(* IEC 61131-3 sources: PLC-IsaVODE/PLC-IsaVODE/samples/plc-programs (part 9) *)

(* ---- 663-GEN_RMP.ST ---- *)
FUNCTION D_TRUNC : DINT
  VAR_INPUT
    x : REAL;
  END_VAR

  D_TRUNC := REAL_TO_DINT(X);
  IF X > 0.0 THEN
  	IF DINT_TO_REAL(D_TRUNC) > X THEN D_TRUNC := D_TRUNC - DINT#1; END_IF;
  ELSE
  	IF DINT_TO_REAL(D_TRUNC) < X THEN D_TRUNC := D_TRUNC + DINT#1; END_IF;
  END_IF;
END_FUNCTION

FUNCTION FRACT:REAL
	VAR_INPUT
		X :	REAL;
	END_VAR

	IF ABS(x) < 2.0E9 THEN
		FRACT := x - DINT_TO_REAL(D_TRUNC(x));
	ELSE
		FRACT := 0.0;
	END_IF;
END_FUNCTION

FUNCTION _REAL_TO_DWORD: DWORD

  VAR_INPUT
    X :	REAL;
  END_VAR

  IF REAL_TO_DWORD(0.5) = DWORD#1 THEN
    _REAL_TO_DWORD := REAL_TO_DWORD(x);
  ELSIF X > 0.0 THEN
    _REAL_TO_DWORD := REAL_TO_DWORD(x+0.5);
  ELSIF X < 0.0 THEN
    _REAL_TO_DWORD := REAL_TO_DWORD(x-0.5);
  ELSE
    _REAL_TO_DWORD := DWORD#0;
  END_IF;
END_FUNCTION

FUNCTION _DWORD_TO_REAL:REAL
	VAR_INPUT
		IN :	DWORD;
	END_VAR

	_DWORD_TO_REAL := UDINT_TO_REAL(DWORD_TO_UDINT(IN));

END_FUNCTION

FUNCTION MULTIME:TIME
	VAR_INPUT
		T :	TIME;
		M :	REAL;
	END_VAR

	multime := DWORD_TO_TIME(_REAL_TO_DWORD(_DWORD_TO_REAL(TIME_TO_DWORD(t))*M));
END_FUNCTION

FUNCTION TIME_TO_REAL1:REAL

VAR_INPUT
	X :	TIME;
END_VAR

TIME_TO_REAL1 := UDINT_TO_REAL(DINT_TO_UDINT(TIME_TO_DINT(X)));
END_FUNCTION

FUNCTION MODR : REAL
  VAR_INPUT
    IN : REAL;
    DIVI : REAL;
  END_VAR

  IF divi = 0.0 THEN
  	MODR := 0.0;
  ELSE
  	MODR := in - DINT_TO_REAL(FLOOR2(in / divi)) * divi;
  END_IF;
END_FUNCTION

FUNCTION FLOOR2 : DINT
  VAR_INPUT
    x : REAL;
  END_VAR

  FLOOR2 := REAL_TO_DINT(X);
  IF DINT_TO_REAL(FLOOR2) > X THEN
  	FLOOR2 := FLOOR2 - DINT#1;
  END_IF;
END_FUNCTION

FUNCTION UDINT_TO_TIME2:TIME

	VAR_INPUT
		IN :	UDINT;
	END_VAR

	UDINT_TO_TIME2 := DINT_TO_TIME(UDINT_TO_DINT(IN));

END_FUNCTION

FUNCTION_BLOCK T_PLC_MS_block
	VAR_OUTPUT
		T_PLC_MS :	UDINT;
	END_VAR

	VAR_EXTERNAL
		PLC_TICKS_PER_SEC :	INT;
		PLC_SYS_TICK_CNT :	DINT;
	END_VAR

	VAR
		debug :	BOOL;(*Debug-Mode ON / OFF*)
		N :	INT;(*Debug-Faktor*)
		Offset :	UDINT;(*Debug-Offset*)
		temp :	DWORD := DWORD#1;(*Debug-Offset*)
		mode :	BOOL;(*modus*)
		faktor :	UDINT;(*Systemtakt-Faktor*)
		init :	BOOL;
		v_plc_ticks_per_sec :	UDINT;
		base :	UDINT := UDINT#1000;
	END_VAR

	IF init = FALSE THEN
		v_plc_ticks_per_sec := INT_TO_UDINT(PLC_TICKS_PER_SEC);
		IF v_plc_ticks_per_sec = UDINT#1024 THEN
			faktor := UDINT#1;
			mode := FALSE;
		ELSIF v_plc_ticks_per_sec > UDINT#0 THEN
			IF v_plc_ticks_per_sec <= base THEN
				faktor := base / v_plc_ticks_per_sec;
				mode := FALSE;
			ELSE
				faktor := v_plc_ticks_per_sec / base;
				mode := TRUE;
			END_IF;
		ELSE
			faktor := UDINT#1;
		END_IF;
		init := TRUE;
	END_IF;

	IF mode THEN
		T_PLC_MS := DINT_TO_UDINT(PLC_SYS_TICK_CNT) / faktor;
	ELSE
		T_PLC_MS := DINT_TO_UDINT(PLC_SYS_TICK_CNT) * faktor;
	END_IF;

	IF debug THEN
		T_PLC_MS := (DWORD_TO_UDINT(SHL(UDINT_TO_DWORD(T_PLC_MS),N) OR SHL(temp,N)) - UDINT#1) + Offset;
	END_IF;

END_FUNCTION_BLOCK

FUNCTION_BLOCK GEN_RMP_Block

	VAR_INPUT
		PT :	TIME := T#1s;
		AM :	REAL := REAL#1.0;
		OS :	REAL;
		DL :	REAL;
	END_VAR

	VAR_OUTPUT
		Q :	BOOL;
		OUT :	REAL;
	END_VAR

	VAR
		tx :	TIME;
		last :	TIME;
		init :	BOOL;
		temp :	REAL;
		ltemp :	REAL;
		T_PLC_MS :	T_PLC_MS_Block;
	END_VAR

	T_PLC_MS();
	tx:= UDINT_TO_TIME(T_PLC_MS.T_PLC_MS) - last;
	DL := modR(dl,1.0);
	IF dl < 0.0 THEN dl := 1.0 - dl; END_IF;

	IF NOT init THEN
		init := TRUE;
		last := tx;
		tx := t#0s;
	END_IF;

	IF tx >= pt THEN
		last := last + pt;
		tx := tx - pt;
	END_IF;

	ltemp := temp;
	IF pt > t#0s THEN temp := fract(TIME_TO_REAL1(tx + multime(pt, dl)) / TIME_TO_REAL1(pt)); END_IF;
	out := am * temp + os;

	Q := temp < ltemp;

END_FUNCTION_BLOCK

PROGRAM program0
  VAR
	PT :	TIME := T#1s;
	AM :	REAL := REAL#1.0;
	OS :	REAL;
	DL :	REAL;
	Q :	BOOL;
	OUT :	REAL;
	func_block : GEN_RMP_Block;
  END_VAR
	func_block.PT  :=PT;
	func_block.AM  :=AM;
	func_block.OS  :=OS;
	func_block.DL  :=DL;
	func_block();
	Q := func_block.Q;
	OUT := func_block.OUT;
END_PROGRAM

CONFIGURATION Config0
	VAR_GLOBAL
		PLC_TICKS_PER_SEC :	INT;
		PLC_SYS_TICK_CNT :	DINT;
	END_VAR
	RESOURCE Res0 ON PLC
		TASK task0(INTERVAL := T#20ms,PRIORITY := 0);
		PROGRAM instance0 WITH task0 : program0;
	END_RESOURCE
END_CONFIGURATION

(* ---- 664-T_AVG24.ST ---- *)
TYPE
  oscat_T_AVG24         	  : ARRAY [0..47]   OF INT;
END_TYPE

FUNCTION_BLOCK T_PLC_MS_block
	VAR_OUTPUT
		T_PLC_MS :	UDINT;
	END_VAR

	VAR_EXTERNAL
		PLC_TICKS_PER_SEC :	INT;
		PLC_SYS_TICK_CNT :	DINT;
	END_VAR

	VAR
		debug :	BOOL;(*Debug-Mode ON / OFF*)
		N :	INT;(*Debug-Faktor*)
		Offset :	UDINT;(*Debug-Offset*)
		temp :	DWORD := DWORD#1;(*Debug-Offset*)
		mode :	BOOL;(*modus*)
		faktor :	UDINT;(*Systemtakt-Faktor*)
		init :	BOOL;
		v_plc_ticks_per_sec :	UDINT;
		base :	UDINT := UDINT#1000;
	END_VAR

	IF init = FALSE THEN
		v_plc_ticks_per_sec := INT_TO_UDINT(PLC_TICKS_PER_SEC);
		IF v_plc_ticks_per_sec = UDINT#1024 THEN
			faktor := UDINT#1;
			mode := FALSE;
		ELSIF v_plc_ticks_per_sec > UDINT#0 THEN
			IF v_plc_ticks_per_sec <= base THEN
				faktor := base / v_plc_ticks_per_sec;
				mode := FALSE;
			ELSE
				faktor := v_plc_ticks_per_sec / base;
				mode := TRUE;
			END_IF;
		ELSE
			faktor := UDINT#1;
		END_IF;
		init := TRUE;
	END_IF;

	IF mode THEN
		T_PLC_MS := DINT_TO_UDINT(PLC_SYS_TICK_CNT) / faktor;
	ELSE
		T_PLC_MS := DINT_TO_UDINT(PLC_SYS_TICK_CNT) * faktor;
	END_IF;

	IF debug THEN
		T_PLC_MS := (DWORD_TO_UDINT(SHL(UDINT_TO_DWORD(T_PLC_MS),N) OR SHL(temp,N)) - UDINT#1) + Offset;
	END_IF;

END_FUNCTION_BLOCK

FUNCTION_BLOCK FILTER_I_Block
	VAR_INPUT
		X :	INT;
		T :	TIME;
	END_VAR

	VAR_OUTPUT
		Y :	INT;
	END_VAR

	VAR
		Yi :	DINT;
		last :	UDINT;
		tx :	UDINT;
		init :	BOOL;
		T_PLC_MS :	T_PLC_MS_block;
	END_VAR

	T_PLC_MS();
	tx:= T_PLC_MS.T_PLC_MS;

	IF NOT init OR T = t#0s THEN
		init := TRUE;
		Yi := INT_TO_DINT(X) * DINT#1000;
	ELSE
		Yi := Yi + INT_TO_DINT(X - Y) * UDINT_TO_DINT(tx - last) * DINT#1000 / TIME_TO_DINT(T);
	END_IF;
	last := tx;
	Y := DINT_TO_INT(yi / DINT#1000);

END_FUNCTION_BLOCK

FUNCTION TIME_TO_UDINT2:UDINT
	VAR_INPUT
		X :	TIME;
	END_VAR

	TIME_TO_UDINT2 := DINT_TO_UDINT(TIME_TO_DINT(X));
END_FUNCTION

FUNCTION INC1:INT

	VAR_INPUT
		X :	INT;
		N :	INT;
	END_VAR

	IF X >= N - 1 THEN
		INC1 := 0;
	ELSE
		INC1 := X + 1;
	END_IF;
END_FUNCTION

FUNCTION_BLOCK T_AVG24_Block

	VAR_INPUT
		TS :	INT;
		DTI :	UDINT;
		RST :	BOOL;
		T_FILTER :	TIME := T#10m;
		SCALE :	REAL := 1.0;
		OFS :	REAL;
	END_VAR

	VAR_OUTPUT
		TA :	REAL;
		_TP :	BOOL;
	END_VAR

	VAR_IN_OUT
		T24 :	REAL;
		T24_MAX :	REAL;
		T24_MIN :	REAL;
	END_VAR

	VAR
		samples :	oscat_T_AVG24;
		pos :	INT;
		init :	BOOL;
		sum :	DINT;
		last :	UDINT;
		tmp_maxxx :	INT;
		tmp_min :	INT;
		i :	INT;
		ft1 :	FILTER_I_Block;
	END_VAR

	ft1(X := TS, T := T_FILTER);

	IF rst OR NOT init THEN
		init := TRUE;
		IF T24 = -1000.0 THEN t24 := INT_TO_REAL(ft1.Y) * 0.1; END_IF;
		FOR pos := 0 TO 47 DO
			samples[pos] := REAL_TO_INT(T24 * 10.0);
		END_FOR;
		pos := 0;
		sum := INT_TO_DINT(samples[0]) * DINT#48;
		TA := (INT_TO_REAL(ft1.Y) * 0.1 + OFS) * SCALE;
		T24 := (DINT_TO_REAL(sum) * 0.00208333333333 + OFS) * SCALE;
		_TP := TRUE;
	ELSIF (dti / UDINT#60 MOD UDINT#30) = UDINT#0 AND DTI > last THEN
		last := DTI + TIME_TO_UDINT2(T#1m);
		sum := sum - INT_TO_DINT(samples[pos]);
		samples[pos] := ft1.Y;
		sum := sum + INT_TO_DINT(samples[pos]);
		pos := INC1(pos, 48);
		TA := (INT_TO_REAL(ft1.Y) * 0.1 + OFS) * SCALE;
		T24 := (DINT_TO_REAL(sum) * 0.00208333333333 + OFS) * SCALE;
		tmp_maxxx := -32000;
		tmp_min := 32000;
		FOR i := 0 TO 47 DO
			tmp_maxxx := MAX(tmp_maxxx, samples[i]);
			tmp_min := MIN(tmp_min, samples[i]);
		END_FOR;
		T24_MAX := (INT_TO_REAL(tmp_maxxx) * 0.1 + OFS) * SCALE;
		T24_MIN := (INT_TO_REAL(tmp_min) * 0.1 + OFS) * SCALE;
		_TP := TRUE;
	ELSE
		_TP := FALSE;
	END_IF;

END_FUNCTION_BLOCK

PROGRAM program0
	VAR
		TS :	INT;
		DTI :	UDINT;
		RST :	BOOL;
		T_FILTER :	TIME := T#10m;
		SCALE :	REAL := 1.0;
		OFS :	REAL;
		TA :	REAL;
		_TP :	BOOL;

		func_block : T_AVG24_Block;
	END_VAR
	func_block.TS := TS;
	func_block.DTI := DTI;
	func_block.RST := RST ;
	func_block.T_FILTER := T_FILTER;
	func_block.SCALE := SCALE;
	func_block.OFS := OFS ;

	func_block();
	TA  := func_block.TA;
	_TP  := func_block._TP;

END_PROGRAM

CONFIGURATION Config0
	VAR_GLOBAL
		PLC_TICKS_PER_SEC :	INT;
		PLC_SYS_TICK_CNT :	DINT;
	END_VAR
  	RESOURCE Res0 ON PLC
    	TASK task0(INTERVAL := T#20ms,PRIORITY := 0);
    	PROGRAM instance0 WITH task0 : program0;
  	END_RESOURCE
END_CONFIGURATION

(* ---- 665-TANK_LEVEL.ST ---- *)
FUNCTION_BLOCK TONOF

	VAR_INPUT
		IN :	BOOL;
		T_ON :	TIME;
		T_OFF :	TIME;
	END_VAR

	VAR_OUTPUT
		Q :	BOOL;
	END_VAR

	VAR
		X :	TON;
		old :	BOOL;
		mode :	BOOL;
	END_VAR

	IF IN XOR old THEN
	X(IN := FALSE, PT := SEL_TIME(IN,T_OFF,T_ON));
	mode := IN;
	old := IN;
	END_IF;
	X(IN := TRUE);
	IF X.Q THEN Q := mode;END_IF;

END_FUNCTION_BLOCK

FUNCTION UDINT_TO_TIME2:TIME

	VAR_INPUT
		IN :	UDINT;
	END_VAR

	UDINT_TO_TIME2 := DINT_TO_TIME(UDINT_TO_DINT(IN));

END_FUNCTION

FUNCTION_BLOCK T_PLC_MS_block
	VAR_OUTPUT
		T_PLC_MS :	UDINT;
	END_VAR

	VAR_EXTERNAL
		PLC_TICKS_PER_SEC :	INT;
		PLC_SYS_TICK_CNT :	DINT;
	END_VAR

	VAR
		debug :	BOOL;(*Debug-Mode ON / OFF*)
		N :	INT;(*Debug-Faktor*)
		Offset :	UDINT;(*Debug-Offset*)
		temp :	DWORD := DWORD#1;(*Debug-Offset*)
		mode :	BOOL;(*modus*)
		faktor :	UDINT;(*Systemtakt-Faktor*)
		init :	BOOL;
		v_plc_ticks_per_sec :	UDINT;
		base :	UDINT := UDINT#1000;
	END_VAR

	IF init = FALSE THEN
		v_plc_ticks_per_sec := INT_TO_UDINT(PLC_TICKS_PER_SEC);
		IF v_plc_ticks_per_sec = UDINT#1024 THEN
			faktor := UDINT#1;
			mode := FALSE;
		ELSIF v_plc_ticks_per_sec > UDINT#0 THEN
			IF v_plc_ticks_per_sec <= base THEN
				faktor := base / v_plc_ticks_per_sec;
				mode := FALSE;
			ELSE
				faktor := v_plc_ticks_per_sec / base;
				mode := TRUE;
			END_IF;
		ELSE
			faktor := UDINT#1;
		END_IF;
		init := TRUE;
	END_IF;

	IF mode THEN
		T_PLC_MS := DINT_TO_UDINT(PLC_SYS_TICK_CNT) / faktor;
	ELSE
		T_PLC_MS := DINT_TO_UDINT(PLC_SYS_TICK_CNT) * faktor;
	END_IF;

	IF debug THEN
		T_PLC_MS := (DWORD_TO_UDINT(SHL(UDINT_TO_DWORD(T_PLC_MS),N) OR SHL(temp,N)) - UDINT#1) + Offset;
	END_IF;
END_FUNCTION_BLOCK

FUNCTION TIME_TO_UDINT2:UDINT
	VAR_INPUT
		X :	TIME;
	END_VAR

	TIME_TO_UDINT2 := DINT_TO_UDINT(TIME_TO_DINT(X));
END_FUNCTION

FUNCTION_BLOCK ACTUATOR_COIL_Block

	VAR_INPUT
		IN :	BOOL;
		SELF_ACT_CYCLE :	TIME := T#10d;
		SELF_ACT_TIME :	TIME := T#1s;
	END_VAR

	VAR_OUTPUT
		OUT :	BOOL;
		STATUS :	BYTE;
	END_VAR

	VAR
		last :	UDINT;
		init :	BOOL;
		tx :	UDINT;
		now :	UDINT;
		T_PLC_MS :	T_PLC_MS_Block;
	END_VAR

	T_PLC_MS();
	now := T_PLC_MS.T_PLC_MS;

	IF NOT init THEN
		last := now;
		init := TRUE;
	ELSIF IN THEN
		OUT := TRUE;
		STATUS := BYTE#101;
		LAST := now;
	ELSE
		OUT := FALSE;
		STATUS := BYTE#100;
		tx := now - last;
		IF (self_act_cycle > T#0s) AND (tx >= TIME_TO_UDINT2(self_act_cycle)) THEN
			OUT := TRUE;
			STATUS := BYTE#102;
			IF tx >= TIME_TO_UDINT2(self_act_cycle + self_act_time) THEN
				last := now;
				OUT := FALSE;
				STATUS := BYTE#100;
			END_IF;
		END_IF;
	END_IF;

END_FUNCTION_BLOCK

FUNCTION_BLOCK TANK_LEVEL_Block

	VAR_INPUT
		LEVEL :	BOOL;
		LEAK :	BOOL;
		ACLR :	BOOL;
		MAX_VALVE_TIME :	TIME;
		LEVEL_DELAY_TIME :	TIME;
	END_VAR

	VAR_OUTPUT
		VALVE :	BOOL;
		ALARM :	BOOL;
		STATUS :	BYTE;
	END_VAR

	VAR
		cx :	ACTUATOR_COIL_Block;
		tn :	TON;
		tl :	TONOF;
		open :	BOOL;
	END_VAR

	tl(in := level, T_ON := level_delay_time, T_OFF := level_delay_time);
	open := tl.Q;

	IF ALARM THEN
		IF ACLR THEN
			ALARM := FALSE;
			STATUS := BYTE#101;
			cx(in := FALSE);
		END_IF;
		RETURN;
	ELSIF LEAK THEN
		cx(in := FALSE);
		ALARM := TRUE;
		STATUS := BYTE#1;
	ELSIF open THEN
		cx(in := TRUE);
		STATUS := BYTE#102;
	ELSE
		cx(in := FALSE);
		STATUS := BYTE#100;
	END_IF;

	tn(in := cx.out AND (MAX_VALVE_TIME > T#0s), PT := MAX_VALVE_TIME);
	IF tn.Q THEN
		ALARM := TRUE;
		STATUS := BYTE#2;
		cx(in := FALSE);
	END_IF;

	VALVE := cx.out;
END_FUNCTION_BLOCK

PROGRAM program0
	VAR
		LEVEL :	BOOL;
		LEAK :	BOOL;
		ACLR :	BOOL;
		MAX_VALVE_TIME :	TIME;
		LEVEL_DELAY_TIME :	TIME;
		VALVE :	BOOL;
		ALARM :	BOOL;
		STATUS :	BYTE;

		func_block : TANK_LEVEL_Block;
	END_VAR
	func_block.LEVEL := LEVEL;
	func_block.LEAK := LEAK;
	func_block.ACLR := ACLR ;
	func_block.MAX_VALVE_TIME := MAX_VALVE_TIME;
	func_block.LEVEL_DELAY_TIME := LEVEL_DELAY_TIME ;
	func_block();
	VALVE  := func_block.VALVE;
	ALARM  := func_block.ALARM;
	STATUS  := func_block.STATUS;
END_PROGRAM

CONFIGURATION Config0
	VAR_GLOBAL
		PLC_TICKS_PER_SEC :	INT;
		PLC_SYS_TICK_CNT :	DINT;
	END_VAR
  	RESOURCE Res0 ON PLC
    	TASK task0(INTERVAL := T#20ms,PRIORITY := 0);
    	PROGRAM instance0 WITH task0 : program0;
  	END_RESOURCE
END_CONFIGURATION

(* ---- 666-M_TX.ST ---- *)
FUNCTION_BLOCK T_PLC_MS_block
	VAR_OUTPUT
		T_PLC_MS :	UDINT;
	END_VAR

	VAR_EXTERNAL
		PLC_TICKS_PER_SEC :	INT;
		PLC_SYS_TICK_CNT :	DINT;
	END_VAR

	VAR
		debug :	BOOL;(*Debug-Mode ON / OFF*)
		N :	INT;(*Debug-Faktor*)
		Offset :	UDINT;(*Debug-Offset*)
		temp :	DWORD := DWORD#1;(*Debug-Offset*)
		mode :	BOOL;(*modus*)
		faktor :	UDINT;(*Systemtakt-Faktor*)
		init :	BOOL;
		v_plc_ticks_per_sec :	UDINT;
		base :	UDINT := UDINT#1000;
	END_VAR

	IF init = FALSE THEN
		v_plc_ticks_per_sec := INT_TO_UDINT(PLC_TICKS_PER_SEC);
		IF v_plc_ticks_per_sec = UDINT#1024 THEN
			faktor := UDINT#1;
			mode := FALSE;
		ELSIF v_plc_ticks_per_sec > UDINT#0 THEN
			IF v_plc_ticks_per_sec <= base THEN
				faktor := base / v_plc_ticks_per_sec;
				mode := FALSE;
			ELSE
				faktor := v_plc_ticks_per_sec / base;
				mode := TRUE;
			END_IF;
		ELSE
			faktor := UDINT#1;
		END_IF;
		init := TRUE;
	END_IF;

	IF mode THEN
		T_PLC_MS := DINT_TO_UDINT(PLC_SYS_TICK_CNT) / faktor;
	ELSE
		T_PLC_MS := DINT_TO_UDINT(PLC_SYS_TICK_CNT) * faktor;
	END_IF;

	IF debug THEN
		T_PLC_MS := (DWORD_TO_UDINT(SHL(UDINT_TO_DWORD(T_PLC_MS),N) OR SHL(temp,N)) - UDINT#1) + Offset;
	END_IF;
END_FUNCTION_BLOCK

FUNCTION_BLOCK M_TX_Block

	VAR_INPUT
		IN :	BOOL;
		TMAX :	TIME := t#10d;
		RST :	BOOL;
	END_VAR

	VAR_OUTPUT
		TH :	TIME;
		TL :	TIME;
		DC :	REAL;
		F :	REAL;
		ET :	TIME;
	END_VAR

	VAR
		edge :	BOOL;
		start :	TIME;
		stop :	TIME;
		tx :	TIME;
		rise :	BOOL;
		fall :	BOOL;
		startup :	BOOL;
		T_PLC_MS :	T_PLC_MS_block;
	END_VAR

	IF rst OR (et >= tmax) THEN
		rise := FALSE;
		fall := FALSE;
		startup := FALSE;
		th := t#0ms;
		tl := t#0ms;
		DC := 0.0;
		F := 0.0;
		ET := t#0s;
	END_IF;

	(* avoid timers to start when input is true at startup *)
	IF NOT startup THEN
		edge := in;
		startup := TRUE;
	END_IF;

	(* read system timer *)
	T_PLC_MS();
	tx:= UDINT_TO_TIME(T_PLC_MS.T_PLC_MS);

	(* edge trigger rising and falling edge *)
	IF in XOR edge THEN
		edge := in;
		(* rising edge starts measurement *)
		IF in THEN
			start := Tx;
			rise := TRUE;
			IF fall THEN tl := start - stop; END_IF;
			IF th > t#0ms AND tl > t#0ms THEN
				dc := TIME_TO_REAL(th) / TIME_TO_REAL(th+tl);
				f := 1000.0 / TIME_TO_REAL(th + tl);
			END_IF;
		(* falling edge starts second cycle measurement *)
		ELSE
			stop := Tx;
			fall := TRUE;
			IF rise THEN th := stop - start; END_IF;
			IF th > t#0ms AND tl > t#0ms THEN
				dc := TIME_TO_REAL(th) /  TIME_TO_REAL(th+tl);
				f := 1000.0 / TIME_TO_REAL(th + tl);
			END_IF;
		END_IF;
	END_IF;
	IF rise THEN et := tx - start; END_IF;

	(* check FOR rst input *)
	IF rst OR (et >= tmax) THEN
		rise := FALSE;
		fall := FALSE;
		startup := FALSE;
		th := t#0ms;
		tl := t#0ms;
		DC := 0.0;
		F := 0.0;
		ET := t#0s;
	END_IF;

	(* avoid timers to start when input is true at startup *)
	IF NOT startup THEN
		edge := in;
		startup := TRUE;
	END_IF;

	(* read system timer *)
	T_PLC_MS();
	tx:= UDINT_TO_TIME(T_PLC_MS.T_PLC_MS);

	(* edge trigger rising and falling edge *)
	IF in XOR edge THEN
		edge := in;
		(* rising edge starts measurement *)
		IF in THEN
			start := Tx;
			rise := TRUE;
			IF fall THEN tl := start - stop; END_IF;
			IF th > t#0ms AND tl > t#0ms THEN
				dc := TIME_TO_REAL(th) / TIME_TO_REAL(th+tl);
				f := 1000.0 / TIME_TO_REAL(th + tl);
			END_IF;
		(* falling edge starts second cycle measurement *)
		ELSE
			stop := Tx;
			fall := TRUE;
			IF rise THEN th := stop - start; END_IF;
			IF th > t#0ms AND tl > t#0ms THEN
				dc := TIME_TO_REAL(th) /  TIME_TO_REAL(th+tl);
				f := 1000.0 / TIME_TO_REAL(th + tl);
			END_IF;
		END_IF;
	END_IF;
	IF rise THEN et := tx - start; END_IF;

END_FUNCTION_BLOCK

PROGRAM program0

	VAR
		IN :	BOOL;
		TMAX :	TIME := t#10d;
		RST :	BOOL;

		TH :	TIME;
		TL :	TIME;
		DC :	REAL;
		F :	REAL;
		ET :	TIME;

		func_block : M_TX_Block;
	END_VAR
	func_block.IN := IN;
	func_block.TMAX := TMAX;
	func_block.RST := RST;

	func_block();
	TH := func_block.TH;
	TL := func_block.TL;
	DC := func_block.DC;
	F := func_block.F;
	ET := func_block.ET;

END_PROGRAM

CONFIGURATION Config0

	VAR_GLOBAL
		PLC_TICKS_PER_SEC :	INT;
		PLC_SYS_TICK_CNT :	DINT;
	END_VAR

	RESOURCE Res0 ON PLC
		TASK task0(INTERVAL := T#20ms,PRIORITY := 0);
		PROGRAM instance0 WITH task0 : program0;
	END_RESOURCE

END_CONFIGURATION

(* ---- 667-METER_STAT.ST ---- *)
FUNCTION DAY_OF_WEEK:INT

	VAR_INPUT
		IDATE :	UDINT;
	END_VAR

	DAY_OF_WEEK := UDINT_TO_INT((idate / UDINT#86400 + UDINT#3) MOD UDINT#7) + INT#01;
END_FUNCTION

FUNCTION LEAP_OF_DATE:BOOL

	VAR_INPUT
		IDATE :	UDINT;
	END_VAR

	LEAP_OF_DATE := SHL(UDINT_TO_DWORD((idate + UDINT#43200) / UDINT#31557600), 30) = DWORD#16#80000000;
END_FUNCTION

FUNCTION DAY_OF_YEAR:INT
	VAR_INPUT
		IDATE :	UDINT;
	END_VAR

	DAY_OF_YEAR := UDINT_TO_INT(((idate) / UDINT#86400) MOD UDINT#1461);
	IF DAY_OF_YEAR > 729 THEN
		IF DAY_OF_YEAR > 1095 THEN DAY_OF_YEAR := DAY_OF_YEAR - 1095; ELSE DAY_OF_YEAR := DAY_OF_YEAR - 729; END_IF;
	ELSIF DAY_OF_YEAR > 364 THEN
		DAY_OF_YEAR := DAY_OF_YEAR - 364;
	ELSE
		DAY_OF_YEAR := DAY_OF_YEAR + 1;
	END_IF;
END_FUNCTION

FUNCTION MONTH_OF_DATE:INT

	VAR_INPUT
		IDATE :	UDINT;
	END_VAR

	MONTH_OF_DATE := DAY_OF_YEAR(idate);
	IF MONTH_OF_DATE < 32 THEN
		MONTH_OF_DATE := 1;
	ELSIF LEAP_OF_DATE((IDATE)) THEN
		MONTH_OF_DATE := (MONTH_OF_DATE * 53 + 1668) / 1623;
	ELSE
		MONTH_OF_DATE := (MONTH_OF_DATE * 53 + 1700) / 1620;
	END_IF;
END_FUNCTION

FUNCTION YEAR_OF_DATE:INT
	VAR_INPUT
		IDATE :	UDINT;
	END_VAR

	YEAR_OF_DATE := UDINT_TO_INT((idate+UDINT#43200) / UDINT#31557600 + UDINT#1970);
END_FUNCTION

FUNCTION_BLOCK METER_STAT_Block

	VAR_INPUT
		IN :	REAL;
		DI :	UDINT;
		RST :	BOOL;
	END_VAR

	VAR_IN_OUT
		LAST_DAY :	REAL;
		CURRENT_DAY :	REAL;
		LAST_WEEK :	REAL;
		CURRENT_WEEK :	REAL;
		LAST_MONTH :	REAL;
		CURRENT_MONTH :	REAL;
		LAST_YEAR :	REAL;
		CURRENT_YEAR :	REAL;
	END_VAR

	VAR RETAIN
		year_start :	REAL;
		month_start :	REAL;
		week_start :	REAL;
		day_start :	REAL;
		last_run :	UDINT;
	END_VAR

	IF rst THEN
		Last_Day := 0.0;
		Current_Day := 0.0;
		Day_start := IN;
		Last_week := 0.0;
		Current_week := 0.0;
		Week_start := in;
		Last_month := 0.0;
		Current_month := 0.0;
		month_start := in;
		last_year := 0.0;
		current_year := 0.0;
		year_start := in;
	ELSE
		Current_Day := IN - Day_Start;
		Current_Week := In - Week_Start;
		Current_Month := IN - Month_Start;
		Current_Year := IN - Year_Start;
	END_IF;

	IF YEAR_OF_DATE(DI) > YEAR_OF_DATE(last_run) THEN
		(* a new year has started *)
		last_year := current_year;
		current_year := 0.0;
		year_start := in;
		last_month := current_month;
		current_month := 0.0;
		month_start := in;
		last_day := current_day;
		current_day := 0.0;
		day_start := in;
	ELSIF MONTH_OF_DATE(DI) > MONTH_OF_DATE(last_run) THEN
		(* a new month has started, january is alrerady done by year change *)
		last_month := current_month;
		current_month := 0.0;
		month_start := in;
		last_day := current_day;
		current_day := 0.0;
		day_start := in;
	ELSIF DAY_OF_YEAR(di) > DAY_OF_YEAR(last_run) THEN
		(* day has chaged, first day of year and first day of month has already been taken care of *)
		last_day := current_day;
		current_day := 0.0;
		day_start := in;
	END_IF;
	IF DAY_OF_WEEK(DI) < DAY_OF_WEEK(last_run) THEN
		(* a new week has started *)
		last_week := current_week;
		current_week := 0.0;
		week_start := in;
	END_IF;
	last_run := di;

END_FUNCTION_BLOCK

PROGRAM program0

	VAR
		IN :	REAL;
		DI :	UDINT;
		RST :	BOOL;

		LAST_DAY :	REAL;
		CURRENT_DAY :	REAL;
		LAST_WEEK :	REAL;
		CURRENT_WEEK :	REAL;
		LAST_MONTH :	REAL;
		CURRENT_MONTH :	REAL;
		LAST_YEAR :	REAL;
		CURRENT_YEAR :	REAL;

		func_block : METER_STAT_Block;
	END_VAR

	func_block.IN := IN;
	func_block.DI := DI;
	func_block.RST := RST;
	func_block.LAST_DAY := LAST_DAY;
	func_block.CURRENT_DAY := CURRENT_DAY;
	func_block.LAST_WEEK := LAST_WEEK;
	func_block.CURRENT_WEEK := CURRENT_WEEK;
	func_block.LAST_MONTH := LAST_MONTH;
	func_block.CURRENT_MONTH := CURRENT_MONTH;
	func_block.LAST_YEAR := LAST_YEAR;
	func_block.CURRENT_YEAR := CURRENT_YEAR;

	func_block();

	LAST_DAY  := func_block.LAST_DAY;
	CURRENT_DAY  := func_block.CURRENT_DAY;
	LAST_WEEK  := func_block.LAST_WEEK;
	CURRENT_WEEK  := func_block.CURRENT_WEEK;
	LAST_MONTH  := func_block.LAST_MONTH;
	CURRENT_MONTH  := func_block.CURRENT_MONTH;
	LAST_YEAR  := func_block.LAST_YEAR;
	CURRENT_YEAR  := func_block.CURRENT_YEAR;

END_PROGRAM

CONFIGURATION Config0

	VAR_GLOBAL
		PLC_TICKS_PER_SEC :	INT;
		PLC_SYS_TICK_CNT :	DINT;
	END_VAR

	RESOURCE Res0 ON PLC
		TASK task0(INTERVAL := T#20ms,PRIORITY := 0);
		PROGRAM instance0 WITH task0 : program0;
	END_RESOURCE

END_CONFIGURATION

(* ---- 668-TN_SC_WRITE_C.ST ---- *)
TYPE
  bya_TN_CHAR:       	ARRAY [0..1919] OF BYTE;
  bya_TN_BACKUP:     	ARRAY [0..1919] OF BYTE;
  bya_TN_COLOR:      	ARRAY [0..1919] OF BYTE;
  bya_TN_Line_Update:	ARRAY [0..23]   OF BOOL;

  us_TN_SCREEN :
  STRUCT
		bya_CHAR:			bya_TN_CHAR;
		bya_COLOR:			bya_TN_COLOR;
		bya_BACKUP:			bya_TN_BACKUP;
		bya_Line_Update:	bya_TN_Line_Update;

		by_Input_Exten_Code:    BYTE;
		by_Input_ASCII_Code:    BYTE;
		bo_Input_ASCII_IsNum:   BOOL;
		in_Page_Number:        	INT;                (* aktive Seiten-Nr.              *)
		in_Cursor_X:           	INT;                (* Cursor X-Position              *)
		in_Cursor_Y:           	INT;                (* Cursor Y-Position              *)
		in_EOS_Offset:         	INT;                (* End of String Offset           *)
		by_Clear_Screen_Attr:  	BYTE;               (* Clear-Screen Attr              *)
		bo_Clear_Screen:       	BOOL;               (* Clear-Screen ausl�sen          *)
		bo_Modal_Dialog:       	BOOL;               (* Modaler Dialog ist aktiv       *)
		bo_Menue_Bar_Dialog:   	BOOL;               (* Menue Dialog ist aktiv         *)

  END_STRUCT;
END_TYPE

FUNCTION _BYTE_TO_INT:INT
	VAR_INPUT
		IN :	BYTE;
	END_VAR

	_BYTE_TO_INT := USINT_TO_INT(BYTE_TO_USINT(IN));
END_FUNCTION

FUNCTION_BLOCK CHR_TO_STRING_Block
	VAR_INPUT
		C :	BYTE;
	END_VAR

	VAR_OUTPUT
		CHR_TO_STRING :	STRING;
	END_VAR

	CHR_TO_STRING := BYTE_TO_STRING(C);

END_FUNCTION_BLOCK

FUNCTION BIT_OF_DWORD : BOOL
  VAR_INPUT
    IN : DWORD;
    N : INT;
  END_VAR

  BIT_OF_DWORD := (SHR(in,N) AND 16#00000001) > 0;
  (* from OSCAT library; www.oscat.de  *)
END_FUNCTION

FUNCTION_BLOCK FILL_Block
	VAR_INPUT
		C :	BYTE;
		L :	INT;
	END_VAR

	VAR_OUTPUT
		FILL :	STRING;
	END_VAR

	VAR
		N :	BYTE;
		I :	INT;
		sx :	STRING;
		CHR_TO_STRING :	CHR_TO_STRING_Block;
		FILL_tmp :	STRING;
	END_VAR

	CHR_TO_STRING(C:=c);
	Sx:=CHR_TO_STRING.CHR_TO_STRING;
	(* create string *)
	N := INT_TO_BYTE(LIMIT(0,L,80));
	(* create a string of characters to be connected to str *)
	FILL := '';
	FOR i := 1 TO 8 DO
		FILL_tmp := FILL;
		FILL := CONCAT(FILL_tmp,FILL);
		IF BIT_OF_DWORD(BYTE_TO_DWORD(N),7) THEN FILL := CONCAT(FILL,Sx); END_IF;
		N := SHL(N,1);
	END_FOR;
END_FUNCTION_BLOCK

FUNCTION_BLOCK FIX_Block

	VAR_INPUT
		STR :	STRING;
		L :	INT;
		C :	BYTE;
		M :	INT;
	END_VAR

	VAR_OUTPUT
		FIX :	STRING;
	END_VAR

	VAR
		N :	INT;
		FILL :	FILL_Block;
	END_VAR

	N := LIMIT(0,L,255) - LEN(str);
	IF N <= 0 THEN
		(* truncate the string at length N *)
		IF M = 1 THEN
			FIX := RIGHT(str,L);
		ELSE
			FIX := LEFT(str,L);
		END_IF;
	ELSIF M = 1 THEN
		(* connect fill characters at the beginning *)
		FILL(C:=C,L:=N);
		FIX := CONCAT(FILL.FILL,str);
	ELSIF M = 2 THEN
		(* center str beween fill characters *)
		(* for an uneven number of fill characters, there is one more at the end *)
		FILL(C:=C,L:=_BYTE_TO_INT(SHR(INT_TO_BYTE(N+1),1)));
		FIX := CONCAT(str,FILL.FILL);
		FILL(C:=C,L:=_BYTE_TO_INT(SHR(INT_TO_BYTE(N),1)));
		FIX := CONCAT(FILL.FILL,FIX);
	ELSE
		(* connect fill characters at the end *)
		FILL(C:=C,L:=N);
		FIX := CONCAT(str,FILL.FILL);
	END_IF;

END_FUNCTION_BLOCK

FUNCTION_BLOCK TN_SC_WRITE_C_Block

	VAR
		FB_FIX :	FIX_Block;
		FB_TN_SC_WRITE :	TN_SC_WRITE;
	END_VAR

	VAR_INPUT
		Iin_Y :	INT;
		Iin_X :	INT;
		Iby_ATTR :	BYTE;
		Ist_STRING :	STRING;
		Iin_LENGTH :	INT;
		Iin_OPTION :	INT;
	END_VAR

	VAR_IN_OUT
		Xus_TN_SCREEN :	us_TN_SCREEN;
	END_VAR

	FB_FIX.str:=Ist_STRING;
	FB_FIX.L:=Iin_LENGTH;
	FB_FIX.C:=BYTE#32;
	FB_FIX.M:=Iin_OPTION;
	FB_FIX();

	FB_TN_SC_WRITE.Iin_Y			:= Iin_Y;
	FB_TN_SC_WRITE.Iin_X			:= Iin_X;
	FB_TN_SC_WRITE.Iby_ATTR			:= Iby_ATTR;
	FB_TN_SC_WRITE.Ist_STRING		:= FB_FIX.FIX;
	FB_TN_SC_WRITE.Xus_TN_SCREEN	:= Xus_TN_SCREEN;
	FB_TN_SC_WRITE();
	Xus_TN_SCREEN := FB_TN_SC_WRITE.Xus_TN_SCREEN;

END_FUNCTION_BLOCK

PROGRAM program0
	VAR
		Iin_Y :	INT;
		Iin_X :	INT;
		Iby_CHAR :	BYTE;
		Xus_TN_SCREEN :	us_TN_SCREEN;

		func_block : TN_SC_WRITE_C_Block;
	END_VAR
	func_block.Iin_Y := Iin_Y;
	func_block.Iin_X := Iin_X;
	func_block.Iby_CHAR := Iby_CHAR;
	func_block.Xus_TN_SCREEN := Xus_TN_SCREEN;

	func_block();
	Xus_TN_SCREEN  := func_block.Xus_TN_SCREEN;
END_PROGRAM

CONFIGURATION Config0
	RESOURCE Res0 ON PLC
		TASK task0(INTERVAL := T#20ms,PRIORITY := 0);
		PROGRAM instance0 WITH task0 : program0;
	END_RESOURCE
END_CONFIGURATION

(* ---- 669-MONTH_TO_STRING.ST ---- *)
TYPE
  oscat_ELEMENT_MONTHS 	: ARRAY [1..12] OF STRING;
  oscat_MONTHS			: ARRAY [1..3]  OF oscat_ELEMENT_MONTHS := [0, 0, 0];
  oscat_ELEMENT_MONTHS3	: ARRAY [1..12] OF STRING;
  oscat_MONTHS3			: ARRAY [1..3]  OF oscat_ELEMENT_MONTHS3 := [0,0,0];
END_TYPE

TYPE oscat_LANGUAGE:
  STRUCT
    DEFAULT 	: INT;
	LMAX    	: INT;
  END_STRUCT;
END_TYPE

FUNCTION_BLOCK SETUP_LANGUAGE_Block

	VAR_IN_OUT
		LANGUAGE :	oscat_LANGUAGE;
	END_VAR

	VAR
		init :	BOOL;
	END_VAR

	IF init THEN RETURN; END_IF;
	init := TRUE;

	LANGUAGE.DEFAULT  := 1; (* 1=english, 2=german 3=french *)
	LANGUAGE.LMAX := 3;
END_FUNCTION_BLOCK

FUNCTION_BLOCK SETUP_MONTHS3_Block

	VAR_IN_OUT
		MONTHS3 :	oscat_MONTHS3;
	END_VAR

	VAR
		init :	BOOL;
	END_VAR

	IF init THEN RETURN; END_IF;
	init := TRUE;

	(* ---- english --- *)
	MONTHS3[1][01] := 'Jan';
	MONTHS3[1][02] := 'Feb';
	MONTHS3[1][03] := 'Mar';
	MONTHS3[1][04] := 'Apr';
	MONTHS3[1][05] := 'May';
	MONTHS3[1][06] := 'Jun';
	MONTHS3[1][07] := 'Jul';
	MONTHS3[1][08] := 'Aug';
	MONTHS3[1][09] := 'Sep';
	MONTHS3[1][10] := 'Oct';
	MONTHS3[1][11] := 'Nov';
	MONTHS3[1][12] := 'Dec';

	(* ---- german --- *)
	MONTHS3[2][01] := 'Jan';
	MONTHS3[2][02] := 'Feb';
	MONTHS3[2][03] := 'Mrz';
	MONTHS3[2][04] := 'Apr';
	MONTHs3[2][05] := 'Mai';
	MONTHS3[2][06] := 'Jun';
	MONTHS3[2][07] := 'Jul';
	MONTHS3[2][08] := 'Aug';
	MONTHS3[2][09] := 'Sep';
	MONTHS3[2][10] := 'Okt';
	MONTHS3[2][11] := 'Nov';
	MONTHS3[2][12] := 'Dez';

	(* ---- french --- *)
	MONTHS3[3][01] := 'Jan';
	MONTHS3[3][02] := 'Fev';
	MONTHS3[3][03] := 'Mar';
	MONTHS3[3][04] := 'Avr';
	MONTHs3[3][05] := 'Mai';
	MONTHS3[3][06] := 'Jun';
	MONTHS3[3][07] := 'Jul';
	MONTHS3[3][08] := 'Aou';
	MONTHS3[3][09] := 'Sep';
	MONTHS3[3][10] := 'Oct';
	MONTHS3[3][11] := 'Nov';
	MONTHS3[3][12] := 'Dec';
	(*@KEY@: END_WORKSHEET *)
END_FUNCTION_BLOCK

FUNCTION_BLOCK SETUP_MONTHS_Block

	VAR_IN_OUT
		MONTHS :	oscat_MONTHS;
	END_VAR

	VAR
		init :	BOOL;
	END_VAR

	IF init THEN RETURN; END_IF;
	init := TRUE;

	(* ---- english --- *)
	MONTHS[1][01] := 'January';
	MONTHS[1][02] := 'February';
	MONTHS[1][03] := 'March';
	MONTHS[1][04] := 'April';
	MONTHS[1][05] := 'May';
	MONTHS[1][06] := 'June';
	MONTHS[1][07] := 'July';
	MONTHS[1][08] := 'August';
	MONTHS[1][09] := 'September';
	MONTHS[1][10] := 'October';
	MONTHS[1][11] := 'November';
	MONTHS[1][12] := 'December';

	(* ---- german --- *)
	MONTHS[2][01] := 'Januar';
	MONTHS[2][02] := 'Februar';
	MONTHS[2][03] := 'March';
	MONTHS[2][04] := 'April';
	MONTHS[2][05] := 'Mai';
	MONTHS[2][06] := 'Juni';
	MONTHS[2][07] := 'Juli';
	MONTHS[2][08] := 'August';
	MONTHS[2][09] := 'September';
	MONTHS[2][10] := 'Oktober';
	MONTHS[2][11] := 'November';
	MONTHS[2][12] := 'Dezember';

	(* ---- french --- *)
	MONTHS[3][01] := 'Janvier';
	MONTHS[3][02] := 'Fvrier';
	MONTHS[3][03] := 'mars';
	MONTHS[3][04] := 'Avril';
	MONTHS[3][05] := 'Mai';
	MONTHS[3][06] := 'Juin';
	MONTHS[3][07] := 'Juillet';
	MONTHS[3][08] := 'Aot';
	MONTHS[3][09] := 'Septembre';
	MONTHS[3][10] := 'Octobre';
	MONTHS[3][11] := 'Novembre';
	MONTHS[3][12] := 'Decembre';
END_FUNCTION_BLOCK

FUNCTION_BLOCK MONTH_TO_STRING_Block

	VAR_INPUT
		MTH :	INT;
		LANG :	INT;
		LX :	INT;
	END_VAR

	VAR_OUTPUT
		MONTH_TO_STRING :	STRING;
	END_VAR

	VAR
		LY :	INT;
		SETUP_MONTHS :	SETUP_MONTHS_Block;
		MONTHS :	oscat_MONTHS;
		SETUP_MONTHS3 :	SETUP_MONTHS3_Block;
		MONTHS3 :	oscat_MONTHS3;
		SETUP_LANGUAGE :	SETUP_LANGUAGE_Block;
		LANGUAGE :	oscat_LANGUAGE;
	END_VAR

	SETUP_MONTHS(MONTHS:=MONTHS);
	MONTHS:=SETUP_MONTHS.MONTHS;
	SETUP_MONTHS3(MONTHS3:=MONTHS3);
	MONTHS3:=SETUP_MONTHS3.MONTHS3;
	SETUP_LANGUAGE(LANGUAGE:=LANGUAGE);
	LANGUAGE:=SETUP_LANGUAGE.LANGUAGE;

	IF LANG = 0 THEN Ly := LANGUAGE.DEFAULT; ELSE ly := MIN(LANG, language.LMAX); END_IF;
	IF MTH < 1 OR MTH > 12 THEN
		RETURN;
	ELSIF LX = 0 THEN
		MONTH_TO_STRING := MONTHS[ly][MTH];
	ELSIF Lx = 3 THEN
		MONTH_TO_STRING := MONTHS3[ly][MTH];
	END_IF;

END_FUNCTION_BLOCK

PROGRAM program0
	VAR
		MTH :	INT;
		LANG :	INT;
		LX :	INT;
		MONTH_TO_STRING :	STRING;
		func_block : MONTH_TO_STRING_Block;
	END_VAR
		func_block.MTH  := MTH;
		func_block.LANG  := LANG;
		func_block.LX  := LX;
		func_block();
		MONTH_TO_STRING := func_block.MONTH_TO_STRING;
END_PROGRAM

CONFIGURATION Config0
	RESOURCE Res0 ON PLC
		TASK task0(INTERVAL := T#20ms,PRIORITY := 0);
		PROGRAM instance0 WITH task0 : program0;
	END_RESOURCE
END_CONFIGURATION

(* ---- 670-WORLD_WEATHER_DESC_GE.ST ---- *)
TYPE
  oscat_STRING3               : STRING;
  oscat_STRING8               : STRING;
  oscat_STRING10              : STRING;
  oscat_STRING60              : STRING;
END_TYPE

TYPE
	oscat_WORLD_WEATHER_CUR :
	STRUCT
		OBSERVATION_TIME : oscat_STRING8;
		TEMP_C           : INT;
		WEATHER_CODE     : INT;
		WEATHER_DESC 	 : oscat_STRING60;
		WEATHER_ICON     : INT;
		WIND_SPEED_MILES : INT;
		WIND_SPEED_KMPH  : INT;
		WIND_DIR_DEGREE  : INT;
		WIND_DIR16POINT  : oscat_STRING3;
		PRECIPMM         : REAL;
		HUMIDITY         : INT;
		VISIBILITY       : INT;
		PRESSURE         : INT;
		CLOUDOVER        : INT;
	END_STRUCT;

	oscat_WORLD_WEATHER_DAY :
	STRUCT
		DATE_OF_DAY      : oscat_STRING10;
		TEMP_MAX_C       : INT;
		TEMP_MAX_F       : INT;
		TEMP_MIN_C       : INT;
		TEMP_MIN_F       : INT;
		WIND_SPEED_MILES : INT;
		WIND_SPEED_KMPH  : INT;
		WIND_DIR_DEGREE  : INT;
		WIND_DIR16POINT  : oscat_STRING3;
		WEATHER_CODE     : INT;
		WEATHER_DESC     : oscat_STRING60;
		WEATHER_ICON     : INT;
		PRECIPMM         : REAL;
	END_STRUCT;

	oscat_WORLD_WEATHER_DAY_ARR : ARRAY [0..4] OF oscat_WORLD_WEATHER_DAY;

	oscat_WORLD_WEATHER_DATA :
	STRUCT
		CUR : oscat_WORLD_WEATHER_CUR;
		DAY : oscat_WORLD_WEATHER_DAY_ARR;
	END_STRUCT;

	oscat_WORLD_WEATHER_aI0_41 : ARRAY[0..41] OF INT;
END_TYPE

FUNCTION_BLOCK WORLD_WEATHER_DESC_GE_Block

	VAR_INPUT
		ACTIVATE :	BOOL;
	END_VAR

	VAR_IN_OUT
		WW :	oscat_WORLD_WEATHER_DATA;
	END_VAR

	VAR
		act_last :	BOOL;
		x :	INT;
		y :	INT;
		str :	oscat_STRING60;
		i :	INT;
	END_VAR

	IF ACTIVATE AND act_last = FALSE THEN
		i := 0;
		FOR y := 1 TO 12 DO
			CASE y OF
			1,3,5,7,9:	x :=  WW.DAY[i].WEATHER_CODE;
			2,4,6,8,10:	WW.DAY[i].WEATHER_DESC := str;
						i := i + 1;
			11:			x :=  WW.CUR.WEATHER_CODE;
			12:			WW.CUR.WEATHER_DESC := str;
			END_CASE;

			CASE x OF
				113	:	str := 'heiter/sonnig';
				116	:	str := 'stellenweise wolkig';
				119	:	str := 'wolkig';
				122	:	str := 'awret';
				143	:	str := 'Nebel';
				176	:	str := 'stellenweise nahegelegener Regen';
				179	:	str := 'stellenweise nahegelegener Schneefall';
				182	:	str := 'stellenweise nahegelegener Eisregen';
				185	:	str := 'stellenweise gefrierender Niesel';
				200	:	str := 'nahegelegene Sturm';
				227	:	str := 'Schneetreiben';
				230	:	str := 'Schneesturm';
				248	:	str := 'Nebel';
				260	:	str := 'gefrierender Nebel';
				263	:	str := 'stellenweise leichter Nieselregen';
				266	:	str := 'leichter Niesel';
				281	:	str := 'gefrierender Nieselregen';
				284	:	str := 'stark gefrierender Nieselregen';
				293	:	str := 'stellenweise leichter Regen';
				296	:	str := 'leichter Regen';
				299	:	str := 'zeitweise etwas Regen';
				302	:	str := 'awerg Regen';
				305	:	str := 'zeitweise etwas starker Regen';
				308	:	str := 'starker Regen';
				311	:	str := 'leichter gefrierender Regen';
				314	:	str := 'awerawer oder starker Eisregen';
				317	:	str := 'leichter Eisregen';
				320	:	str := 'awewea oder starker Eisregen';
				323	:	str := 'stellenweise leichter Schneefall';
				326	:	str := 'leichter Scheefall';
				329	:	str := 'stellenweise moderater Schneefall';
				332	:	str := 'awertwy Schnee';
				335	:	str := 'stellenweise starker Scheefall';
				338	:	str := 'starker Schneefall';
				350	:	str := 'Hagel';
				353	:	str := 'leichte ewruerh';
				356	:	str := 'awerwaer oder starker Regenfall';
				359	:	str := 'sintflutartige aweheawh';
				362	:	str := 'leichter Eisregen';
				365	:	str := 'aweraweb oder starker Eisregen';
				368	:	str := 'leichte Schneeschauer';
				371	:	str := 'awerawb oder starker Schneefall';
				374	:	str := 'leichter Hagel';
				377	:	str := 'awerawer oder starker Hagel';
				386	:	str := 'stellenweise leichter Regen in Gewittergebiet';
				389	:	str := 'awer oder starker Regen in Gewittergebiet';
				392	:	str := 'stellenweise leichter Schneefall in Gewittergebiet';
				395	:	str := 'awerh oder starker Schnee in Gewittergebiet';
			ELSE
				str := 	'nicht aweh';
			END_CASE;
		END_FOR;
	END_IF;
	act_last := ACTIVATE;

END_FUNCTION_BLOCK

PROGRAM program0
	VAR
		ACTIVATE :	BOOL;
		WW :	oscat_WORLD_WEATHER_DATA;

		func_block : WORLD_WEATHER_DESC_GE_Block;
	END_VAR
	func_block.ACTIVATE := ACTIVATE;
	func_block.WW := WW;

	func_block();
	WW  := func_block.WW;
END_PROGRAM

CONFIGURATION Config0
	RESOURCE Res0 ON PLC
		TASK task0(INTERVAL := T#20ms,PRIORITY := 0);
		PROGRAM instance0 WITH task0 : program0;
	END_RESOURCE
END_CONFIGURATION

(* ---- 671-LOG_VIEWPORT.ST ---- *)
TYPE
  oscat_STRING80             : STRING;
  oscat_STRING250             : STRING;
END_TYPE

TYPE
  PRINTF_DATA_250  	:  ARRAY [1..11]  OF oscat_STRING250;
  PRINTF_DATA_80 	:  ARRAY [1..11]  OF oscat_STRING80;
  LOG_250       	:  ARRAY [0..400] OF oscat_STRING250;
  LOG_80    		:  ARRAY [0..400] OF oscat_STRING80;
  LOG_OPTION		:  ARRAY [0..400] OF DWORD;

  us_LOG_CONTROL :
  STRUCT
    NEW_MSG              : oscat_STRING250;    (*W neue Nachricht f�r den Datenbuffer   *)
	NEW_MSG_OPTION 		 : DWORD;
    LEVEL                : BYTE;
	SIZE                 : INT;                (*R Anzahl der Strings im LOG_DATA       *)
	RESET                : BOOL;               (*W Nachrichtenbuffer l�schen            *)
    PRINTF               : PRINTF_DATA_250;    (*W Array PRINTF Parameter               *)
    MSG                  : LOG_250;            (*I Array Message                        *)
    MSG_OPTION           : LOG_OPTION;     	   (*I Array Message Option                 *)
	UPDATE_COUNT         : UINT;               (*R Updatez�hler                         *)
    IDX                  : INT;                (*R aktueller Nachrichten-Index          *)
	RING_MODE            : BOOL;               (*I Buffer�berlauf erkannt               *)
  END_STRUCT;

  us_LOG_CONTROL_80 :
  STRUCT
    NEW_MSG              : oscat_STRING80;     (*W neue Nachricht f�r den Datenbuffer   *)
	NEW_MSG_OPTION 		 : DWORD;
    LEVEL                : BYTE;
	SIZE                 : INT;                (*R Anzahl der Strings im LOG_DATA       *)
	RESET                : BOOL;               (*W Nachrichtenbuffer l�schen            *)
    PRINTF               : PRINTF_DATA_80;     (*W Array PRINTF Parameter               *)
    MSG                  : LOG_80;             (*I Array Message                        *)
    MSG_OPTION           : LOG_OPTION;     	   (*I Array Message Option                 *)
	UPDATE_COUNT         : UINT;               (*R Updatez�hler                         *)
    IDX                  : INT;                (*R aktueller Nachrichten-Index          *)
	RING_MODE            : BOOL;               (*I Buffer�berlauf erkannt               *)
  END_STRUCT;

  LINE_ARRAY 			: ARRAY [1..40] OF INT;

  us_LOG_VIEWPORT :
    STRUCT
     LINE_ARRAY          : LINE_ARRAY;
     COUNT               : INT;                (* Anzahl der sichtbaren Nachtrichten   *)
	 UPDATE_COUNT        : UINT;               (* Updatez�hler                         *)
     MOVE_TO_X           : INT;                (* Steuerung der Nachrichtenanzeige     *)
     UPDATE              : BOOL;               (* Daten wurden ge�ndert -> neuzeichnen *)
  END_STRUCT;

END_TYPE

FUNCTION_BLOCK LOG_VIEWPORT_Block

  VAR_IN_OUT
    LC :	us_LOG_CONTROL_80;
    LV :	us_LOG_VIEWPORT;
  END_VAR

  VAR
    pos :	INT;
    count :	INT;
    idx :	INT;
    base :	INT;
    update_pos :	BOOL;
  END_VAR

  IF LV.MOVE_TO_X <> 0 THEN
    CASE LV.MOVE_TO_X OF
    30000:
      pos := 1 ;
    30001:
      pos := LC.SIZE;
    30002:
      pos := pos + LV.COUNT;
    30003:
      pos := pos - LV.COUNT;
    ELSE
      pos := pos + LV.MOVE_TO_X;
    END_CASE;
    update_pos := TRUE;
    LV.MOVE_TO_X := 0;
  END_IF;

  IF (LV.UPDATE_COUNT <> LC.UPDATE_COUNT) OR update_pos THEN
    LV.UPDATE := TRUE;
    LV.UPDATE_COUNT := LC.UPDATE_COUNT;
    update_pos := FALSE;

    IF LC.RING_MODE THEN
      pos := LIMIT(1,pos,LC.SIZE - LV.COUNT + 1);
    ELSE
      IF LC.IDX > LV.COUNT THEN
        pos := LIMIT(1,pos,LC.IDX - LV.COUNT + 1);
      ELSE
        pos := 1;
      END_IF;
    END_IF;

    base := LC.IDX - pos - LV.COUNT + 1;
    IF LC.RING_MODE THEN
      FOR count:= 1 TO LV.COUNT DO
        idx := base + count;
        IF idx < 1 THEN
          idx := idx + LC.SIZE;
        END_IF;
      END_FOR;
    ELSE
      FOR count:= 1 TO LV.COUNT DO
        idx := base + count;
        IF idx < 1 THEN
          LV.LINE_ARRAY[count] := 0;
        ELSE
          LV.LINE_ARRAY[count] := idx;
        END_IF;
      END_FOR;
    END_IF;
  END_IF;

END_FUNCTION_BLOCK

PROGRAM program0
	VAR
		LC :	us_LOG_CONTROL_80;
    LV :	us_LOG_VIEWPORT;

		func_block : LOG_VIEWPORT_Block;
	END_VAR
	func_block.LC := LC;
	func_block.LV := LV;

	func_block();
  LC  := func_block.LC;
  LV  := func_block.LV;

END_PROGRAM

CONFIGURATION Config0

  	RESOURCE Res0 ON PLC
    	TASK task0(INTERVAL := T#20ms,PRIORITY := 0);
    	PROGRAM instance0 WITH task0 : program0;
  	END_RESOURCE

END_CONFIGURATION

(* ---- 672-CTRL_PI.ST ---- *)
FUNCTION_BLOCK T_PLC_US_Block
	VAR_OUTPUT
		T_PLC_US :	UDINT;
	END_VAR

	VAR_EXTERNAL
		PLC_TICKS_PER_SEC :	INT;
		PLC_SYS_TICK_CNT :	DINT;
	END_VAR

	VAR
		debug :	BOOL;
		N :	INT;
		Offset :	UDINT;
		temp :	DWORD := DWORD#1;
		mode :	BOOL;
		faktor :	UDINT;
		init :	BOOL;
		v_plc_ticks_per_sec :	UDINT;
		base :	UDINT := UDINT#1000000;
	END_VAR

	IF init = FALSE THEN
		v_plc_ticks_per_sec := INT_TO_UDINT(PLC_TICKS_PER_SEC);
		IF v_plc_ticks_per_sec = UDINT#1024 THEN
			faktor := UDINT#1000;
			mode := FALSE;
		ELSIF v_plc_ticks_per_sec > UDINT#0 THEN
			IF v_plc_ticks_per_sec <= base THEN
				faktor := base / v_plc_ticks_per_sec;
				mode := FALSE;
			ELSE
				faktor := v_plc_ticks_per_sec / base;
				mode := TRUE;
			END_IF;
		ELSE
			faktor := UDINT#1;
		END_IF;
		init := TRUE;
	END_IF;

	IF mode THEN
		T_PLC_US := DINT_TO_UDINT(PLC_SYS_TICK_CNT) / faktor;
	ELSE
		T_PLC_US := DINT_TO_UDINT(PLC_SYS_TICK_CNT) * faktor;
	END_IF;

	IF debug THEN
		T_PLC_US := (DWORD_TO_UDINT(SHL(UDINT_TO_DWORD(T_PLC_US),N) OR SHL(temp,N)) - UDINT#1) + Offset;
	END_IF;
END_FUNCTION_BLOCK

FUNCTION_BLOCK FT_PIWL

	VAR_INPUT
		IN :	REAL;
		KP :	REAL := 1.0;
		KI :	REAL := 1.0;
		LIM_L :	REAL := -1.0E38;
		LIM_H :	REAL := 1.0E38;
		RST :	BOOL;
	END_VAR

	VAR_OUTPUT
		Y :	REAL;
		LIM :	BOOL;
	END_VAR

	VAR
		init :	BOOL;
		tx :	UDINT;
		tc :	REAL;
		t_last :	UDINT;
		in_last :	REAL;
		i :	REAL;
		p :	REAL;
		T_PLC_US :	T_PLC_US_Block;
	END_VAR

	IF NOT init OR RST THEN
		init := TRUE;
		in_last := in;
		T_PLC_US();
		t_last := T_PLC_US.T_PLC_US;
		i := 0.0;
		tc := 0.0;
	ELSE
		(* read last cycle time in Microseconds *)
		T_PLC_US();
		tx := T_PLC_US.T_PLC_US;
		tc := UDINT_TO_REAL(tx - t_last);
		t_last := tx;

		(* calculate proportional part *)
		p := KP * IN;

		(* run integrator *)
		i := (IN + in_last) * 5.0E-7 * KI * tc + i;
		in_last := IN;

		(* calculate output Y *)
		Y := p + i;

		(* check output for limits *)
		IF Y >= LIM_H THEN
			Y := LIM_H;
			IF ki <> 0.0 THEN
				i := LIM_H - p;
			ELSE
				i := 0.0;
			END_IF;
			LIM := TRUE;
		ELSIF Y <= LIM_L THEN
			Y := LIM_L;
			IF ki <> 0.0 THEN
				i := LIM_L - p;
			ELSE
				i := 0.0;
			END_IF;
			LIM := TRUE;
		ELSE
			LIM := FALSE;
		END_IF;
	END_IF;
END_FUNCTION_BLOCK

FUNCTION_BLOCK CTRL_OUT
	VAR_INPUT
		CI :	REAL;
		OFFSET :	REAL;
		MAN_IN :	REAL;
		LIM_L :	REAL;
		LIM_H :	REAL;
		MANUAL :	BOOL;
	END_VAR

	VAR_OUTPUT
		Y :	REAL;
		LIM :	BOOL;
	END_VAR

	Y := SEL(manual, CI, MAN_IN) + OFFSET;

	IF Y >= LIM_H THEN
		Y := LIM_H;
		LIM := TRUE;
	ELSIF Y <= lim_L THEN
		Y := LIM_L;
		LIM := TRUE;
	ELSE
		LIM := FALSE;
	END_IF;
END_FUNCTION_BLOCK

FUNCTION DEAD_ZONE:REAL

	VAR_INPUT
		X :	REAL;
		L :	REAL;
	END_VAR

	IF ABS(x) > L THEN
		dead_zone := X;
	ELSE
		DEAD_ZONE := 0.0;
	END_IF;

END_FUNCTION

FUNCTION CTRL_IN:REAL
	VAR_INPUT
		SET_POINT :	REAL;
		ACTUAL :	REAL;
		NOISE :	REAL;
	END_VAR
	CTRL_IN := DEAD_ZONE(SET_POINT - ACTUAL, NOISE);
END_FUNCTION

FUNCTION_BLOCK CTRL_PI
	VAR_INPUT
		ACT :	REAL;
		SET :	REAL;
		SUP :	REAL;
		OFS :	REAL;
		M_I :	REAL;
		MAN :	BOOL;
		RST :	BOOL := FALSE;
		KP  :	REAL := 1.0;
		KI  :	REAL := 1.0;
		LL  :	REAL := -1000.0;
		LH  :	REAL := 1000.0;
	END_VAR

	VAR_OUTPUT
		Y    :	REAL;
		DIFF :	REAL;
		LIM  :	BOOL;
	END_VAR

	VAR
		pi :	FT_PIWL;
		co :	CTRL_OUT;
	END_VAR

	DIFF := CTRL_IN(SET, ACT, SUP);
	pi(in := DIFF, kp := KP, ki := KI, lim_l := LL, lim_h := LH, rst := RST);
	co(ci := pi.Y, OFFSET := OFS, man_in := M_I, lim_l := LL, lim_h := LH, manual := MAN);
	Y := co.Y;
	LIM := co.LIM;
END_FUNCTION_BLOCK

PROGRAM program0
  VAR
		ACT :	REAL;
		SET :	REAL;
		SUP :	REAL;
		OFS :	REAL;
		M_I :	REAL;
		MAN :	BOOL;
		RST :	BOOL;
		KP  :	REAL;
		KI  :	REAL;
		LL  :	REAL;
		LH  :	REAL;

		Y    :	REAL;
		DIFF :	REAL;
		LIM  :	BOOL;

	func_block : CTRL_PI;
  END_VAR
	func_block.ACT  :=ACT ;
	func_block.SET  :=SET ;
	func_block.SUP  :=SUP ;
	func_block.OFS  :=OFS ;
	func_block.M_I  :=M_I ;
	func_block.MAN  :=MAN ;
	func_block.RST  :=RST ;
	func_block.KP   :=KP  ;
	func_block.KI   :=KI  ;
	func_block.LL   :=LL  ;
	func_block.LH   :=LH  ;

	func_block();
	Y    := func_block.Y   ;
	DIFF := func_block.DIFF;
	LIM  := func_block.LIM ;
END_PROGRAM

CONFIGURATION Config0
	VAR_GLOBAL
		PLC_TICKS_PER_SEC :	INT;
		PLC_SYS_TICK_CNT :	DINT;
	END_VAR

	RESOURCE Res0 ON PLC
		TASK task0(INTERVAL := T#20ms,PRIORITY := 0);
		PROGRAM instance0 WITH task0 : program0;
	END_RESOURCE
END_CONFIGURATION

(* ---- 673-FT_PIDWL.ST ---- *)
FUNCTION_BLOCK T_PLC_US_Block
	VAR_OUTPUT
		T_PLC_US :	UDINT;
	END_VAR

	VAR_EXTERNAL
		PLC_TICKS_PER_SEC :	INT;
		PLC_SYS_TICK_CNT :	DINT;
	END_VAR

	VAR
		debug :	BOOL;
		N :	INT;
		Offset :	UDINT;
		temp :	DWORD := DWORD#1;
		mode :	BOOL;
		faktor :	UDINT;
		init :	BOOL;
		v_plc_ticks_per_sec :	UDINT;
		base :	UDINT := UDINT#1000000;
	END_VAR

	IF init = FALSE THEN
		v_plc_ticks_per_sec := INT_TO_UDINT(PLC_TICKS_PER_SEC);
		IF v_plc_ticks_per_sec = UDINT#1024 THEN
			faktor := UDINT#1000;
			mode := FALSE;
		ELSIF v_plc_ticks_per_sec > UDINT#0 THEN
			IF v_plc_ticks_per_sec <= base THEN
				faktor := base / v_plc_ticks_per_sec;
				mode := FALSE;
			ELSE
				faktor := v_plc_ticks_per_sec / base;
				mode := TRUE;
			END_IF;
		ELSE
			faktor := UDINT#1;
		END_IF;
		init := TRUE;
	END_IF;

	IF mode THEN
		T_PLC_US := DINT_TO_UDINT(PLC_SYS_TICK_CNT) / faktor;
	ELSE
		T_PLC_US := DINT_TO_UDINT(PLC_SYS_TICK_CNT) * faktor;
	END_IF;

	IF debug THEN
		T_PLC_US := (DWORD_TO_UDINT(SHL(UDINT_TO_DWORD(T_PLC_US),N) OR SHL(temp,N)) - UDINT#1) + Offset;
	END_IF;
END_FUNCTION_BLOCK

FUNCTION_BLOCK FT_PIWL

	VAR_INPUT
		IN :	REAL;
		KP :	REAL := 1.0;
		KI :	REAL := 1.0;
		LIM_L :	REAL := -1.0E38;
		LIM_H :	REAL := 1.0E38;
		RST :	BOOL;
	END_VAR

	VAR_OUTPUT
		Y :	REAL;
		LIM :	BOOL;
	END_VAR

	VAR
		init :	BOOL;
		tx :	UDINT;
		tc :	REAL;
		t_last :	UDINT;
		in_last :	REAL;
		i :	REAL;
		p :	REAL;
		T_PLC_US :	T_PLC_US_Block;
	END_VAR

	IF NOT init OR RST THEN
		init := TRUE;
		in_last := in;
		T_PLC_US();
		t_last := T_PLC_US.T_PLC_US;
		i := 0.0;
		tc := 0.0;
	ELSE
		(* read last cycle time in Microseconds *)
		T_PLC_US();
		tx := T_PLC_US.T_PLC_US;
		tc := UDINT_TO_REAL(tx - t_last);
		t_last := tx;

		(* calculate proportional part *)
		p := KP * IN;

		(* run integrator *)
		i := (IN + in_last) * 5.0E-7 * KI * tc + i;
		in_last := IN;

		(* calculate output Y *)
		Y := p + i;

		(* check output for limits *)
		IF Y >= LIM_H THEN
			Y := LIM_H;
			IF ki <> 0.0 THEN
				i := LIM_H - p;
			ELSE
				i := 0.0;
			END_IF;
			LIM := TRUE;
		ELSIF Y <= LIM_L THEN
			Y := LIM_L;
			IF ki <> 0.0 THEN
				i := LIM_L - p;
			ELSE
				i := 0.0;
			END_IF;
			LIM := TRUE;
		ELSE
			LIM := FALSE;
		END_IF;
	END_IF;
END_FUNCTION_BLOCK

FUNCTION_BLOCK FT_DERIV
	VAR_INPUT
		IN :	REAL;
		K :	REAL := 1.0;
		RUN :	BOOL := TRUE;
	END_VAR

	VAR_OUTPUT
		OUT :	REAL;
	END_VAR

	VAR
		old :	REAL;
		tx :	UDINT;
		last :	UDINT;
		init :	BOOL;
		tc :	REAL;
		T_PLC_US :	T_PLC_US_Block;
	END_VAR

	T_PLC_US();
	tx:= T_PLC_US.T_PLC_US;
	tc := UDINT_TO_REAL(tx - last);

	IF NOT init THEN
		init := TRUE;
		old := in;
	ELSIF run AND tc > 0.0 THEN
		out := (in - old) / tc * 1000000.0 * K;
		old := in;
	ELSE
		out := 0.0;
	END_IF;

	last := tx;

	T_PLC_US();
	tx:= T_PLC_US.T_PLC_US;

	IF NOT init THEN
		init := TRUE;
	ELSIF run AND tx - last > UDINT#0 THEN
		out := (in - old) / UDINT_TO_REAL(tx - last) * 1000000.0 * K;
	ELSE
		out := 0.0;
	END_IF;
	old := in;
	last := tx;
END_FUNCTION_BLOCK

FUNCTION_BLOCK FT_PIDWL
	VAR_INPUT
		IN :	REAL;
		KP :	REAL := 1.0;
		TN :	REAL := 1.0;
		TV :	REAL := 1.0;
		LIM_L :	REAL := -1.0E38;
		LIM_H :	REAL := 1.0E38;
		RST :	BOOL;
	END_VAR

	VAR_OUTPUT
		Y :	REAL;
		LIM :	BOOL;
	END_VAR

	VAR
		piwl :	FT_PIWL;
		diff :	FT_DERIV;
	END_VAR

	IF rst THEN
		piwl(rst := TRUE);
		piwl.RST := FALSE;
	ELSE
		IF TN = 0.0 THEN
			piwl(in := IN * KP, KP := 1.0, KI := 0.0, LIM_L := LIM_L, LIM_H := LIM_H);
		ELSE
			piwl(in := IN * KP, KP := 1.0, KI := 1.0 / TN, LIM_L := LIM_L, LIM_H := LIM_H);
		END_IF;

		diff(IN := IN, K := KP * TV);
		Y := piwl.Y + diff.out;

		IF Y < LIM_L THEN
			LIM := TRUE;
			Y := LIM_L;
		ELSIF Y > LIM_H THEN
			LIM := TRUE;
			Y := LIM_H;
		ELSE
			LIM := FALSE;
		END_IF;
	END_IF;
END_FUNCTION_BLOCK

PROGRAM program0
  VAR
	IN    :	REAL;
	KP    :	REAL;
	TN    :	REAL;
	TV    :	REAL;
	LIM_L :	REAL;
	LIM_H :	REAL;
	RST   :	BOOL;

	Y :	REAL;
	LIM :	BOOL;

	func_block : FT_PIDWL;
  END_VAR
	func_block.IN    :=IN   ;
	func_block.KP    :=KP   ;
	func_block.TN    :=TN   ;
	func_block.TV    :=TV   ;
	func_block.LIM_L :=LIM_L;
	func_block.LIM_H :=LIM_H;
	func_block.RST   :=RST  ;
	func_block();
	Y := func_block.Y;
	LIM := func_block.LIM;
END_PROGRAM

CONFIGURATION Config0
	VAR_GLOBAL
		PLC_TICKS_PER_SEC :	INT;
		PLC_SYS_TICK_CNT :	DINT;
	END_VAR

	RESOURCE Res0 ON PLC
		TASK task0(INTERVAL := T#20ms,PRIORITY := 0);
		PROGRAM instance0 WITH task0 : program0;
	END_RESOURCE
END_CONFIGURATION

(* ---- 674-MATRIX.ST ---- *)
TYPE
	oscat_arb_0_3               : ARRAY [0..3]    OF BYTE;
END_TYPE

FUNCTION BIT_OF_DWORD : BOOL
	VAR_INPUT
		IN : DWORD;
		N : INT;
	END_VAR

	BIT_OF_DWORD := (SHR(in,N) AND 16#00000001) > 0;
END_FUNCTION

FUNCTION _BYTE_TO_INT:INT
	VAR_INPUT
		IN :	BYTE;
	END_VAR

	_BYTE_TO_INT := USINT_TO_INT(BYTE_TO_USINT(IN));
END_FUNCTION

FUNCTION BIT_LOAD_B:BYTE
	VAR_INPUT
		IN :	BYTE;
		VAL :	BOOL;
		POS :	INT;
	END_VAR

	IF VAL THEN
		BIT_LOAD_B := in OR SHL(BYTE#1,pos);
	ELSE
		BIT_LOAD_B := in AND (NOT SHL(BYTE#1,pos));
	END_IF;
END_FUNCTION

FUNCTION_BLOCK MATRIX_Block

	VAR_INPUT
		X1 :	BOOL;
		X2 :	BOOL;
		X3 :	BOOL;
		X4 :	BOOL;
		X5 :	BOOL;
		RELEASE :	BOOL;
	END_VAR

	VAR_OUTPUT
		CODE :	BYTE;
		_TP :	BOOL;
		Y1 :	BOOL := TRUE;
		Y2 :	BOOL;
		Y3 :	BOOL;
		Y4 :	BOOL;
	END_VAR

	VAR
		line :	BYTE;
		X :	oscat_arb_0_3;
		L :	oscat_arb_0_3;
		i :	INT;
		temp :	BYTE;
		temp2 :	BYTE;
		L_temp :	BYTE;
		temp_bit :	BOOL;
		in_temp :	INT;
	END_VAR

	_TP := FALSE;
	code := BYTE#0;

	(* read scan lines *)
	in_temp := _BYTE_TO_INT(line);
	temp := X[in_temp];  (* X[LINE] umkopieren *)

	temp:=BIT_LOAD_B(temp,X1,0); (* X[line].0 := X1; *)
	temp:=BIT_LOAD_B(temp,X2,1); (* X[line].1 := X2; *)
	temp:=BIT_LOAD_B(temp,X3,2); (* X[line].2 := X3; *)
	temp:=BIT_LOAD_B(temp,X4,3); (* X[line].3 := X4; *)
	temp:=BIT_LOAD_B(temp,X5,4); (* X[line].4 := X5; *)

	X[in_temp] := temp; (* X[LINE] zur�ckkopieren *)

	(* compare for change *)
	FOR i := 0 TO 3 DO
		IF X[i] <> L[i] THEN
			(* scan line information has changed code need to be found and generated *)
			temp   := x[i] XOR L[i];
			temp2  := X[i];
			L_temp := L[i];

			IF BIT_OF_DWORD(BYTE_TO_DWORD(temp),0) THEN (* temp.X0 *)
				code := BYTE#1;
				temp_bit := BIT_OF_DWORD(BYTE_TO_DWORD(temp2),0);   (* X[i].X0 *)
				code := BIT_LOAD_B(code,temp_bit,7);     			(* code.X7 *)
				L_temp := BIT_LOAD_B(L_temp,temp_bit,0); 			(* L[i].X0 *)
			ELSIF BIT_OF_DWORD(BYTE_TO_DWORD(temp),1) THEN          (* temp.X1 *)
				code := BYTE#2;
				temp_bit := BIT_OF_DWORD(BYTE_TO_DWORD(temp2),1);   (* X[i].X1 *)
				code := BIT_LOAD_B(code,temp_bit,7);     			(* code.X7 *)
				L_temp := BIT_LOAD_B(L_temp,temp_bit,1); 			(* L[i].X1 *)
			ELSIF BIT_OF_DWORD(BYTE_TO_DWORD(temp),2) THEN          (* temp.X2 *)
				code := BYTE#3;
				temp_bit := BIT_OF_DWORD(BYTE_TO_DWORD(temp2),2);   (* X[i].X2 *)
				code := BIT_LOAD_B(code,temp_bit,7);     			(* code.X7 *)
				L_temp := BIT_LOAD_B(L_temp,temp_bit,2); 			(* L[i].X2 *)
			ELSIF BIT_OF_DWORD(BYTE_TO_DWORD(temp),3) THEN          (* temp.X3 *)
				code := BYTE#4;
				temp_bit := BIT_OF_DWORD(BYTE_TO_DWORD(temp2),3);   (* X[i].X3 *)
				code := BIT_LOAD_B(code,temp_bit,7);     			(* code.X7 *)
				L_temp := BIT_LOAD_B(L_temp,temp_bit,3); 			(* L[i].X3 *)
			ELSIF BIT_OF_DWORD(BYTE_TO_DWORD(temp),4) THEN          (* temp.X4 *)
				code := BYTE#5;
				temp_bit := BIT_OF_DWORD(BYTE_TO_DWORD(temp2),4);   (* X[i].X4 *)
				code := BIT_LOAD_B(code,temp_bit,7);     			(* code.X7 *)
				L_temp := BIT_LOAD_B(L_temp,temp_bit,4); 			(* L[i].X4 *)
			END_IF;
			L[i] := L_temp;
			_TP := TRUE;
			code := (code AND BYTE#2#1000_1111) OR SHL(LINE AND BYTE#2#0000_0111,4);
			(* obere zeile enspricht: Code.X4 := Line.X0; /  Code.X5 := Line.X1; / Code.X6 := Line.X2; *)

			(* check if release codes need to be killed *)
			IF NOT release AND code < BYTE#127 THEN
				code := BYTE#0;
				_TP := FALSE;
			END_IF;
			EXIT;
		END_IF;
	END_FOR;

	(* increment scan line every cycle *)
	line := INT_TO_BYTE(_BYTE_TO_INT(line) + 1) AND BYTE#2#0000_0011;
	temp := SHL(BYTE#1,_BYTE_TO_INT(line));

	Y1 := BIT_OF_DWORD(BYTE_TO_DWORD(temp),0); (* temp.0 *)
	Y2 := BIT_OF_DWORD(BYTE_TO_DWORD(temp),1); (* temp.1 *)
	Y3 := BIT_OF_DWORD(BYTE_TO_DWORD(temp),2); (* temp.2 *)
	Y4 := BIT_OF_DWORD(BYTE_TO_DWORD(temp),3); (* temp.3 *)

END_FUNCTION_BLOCK

PROGRAM program0

	VAR
		X1 :	BOOL;
		X2 :	BOOL;
		X3 :	BOOL;
		X4 :	BOOL;
		X5 :	BOOL;
		RELEASE :	BOOL;

		CODE :	BYTE;
		_TP :	BOOL;
		Y1 :	BOOL := TRUE;
		Y2 :	BOOL;
		Y3 :	BOOL;
		Y4 :	BOOL;

		func_block : MATRIX_Block;
	END_VAR
	func_block.X1 := X1;
	func_block.X2 := X2;
	func_block.X3 := X3;
	func_block.X4 := X4;
	func_block.X5 := X5;
	func_block.RELEASE := RELEASE;
	func_block();
	CODE := func_block.CODE;
	_TP := func_block._TP;
	Y1 := func_block.Y1;
	Y2 := func_block.Y2;
	Y3 := func_block.Y3;
	Y4 := func_block.Y4;

END_PROGRAM

CONFIGURATION Config0

	RESOURCE Res0 ON PLC
		TASK task0(INTERVAL := T#20ms,PRIORITY := 0);
		PROGRAM instance0 WITH task0 : program0;
	END_RESOURCE

END_CONFIGURATION

(* ---- 675-TN_INPUT_SELECT_POPUP.ST ---- *)
FUNCTION_BLOCK TN_INPUT_SELECT_POPUP

  VAR
    in_index :	INT;
    in_Element_Count :	INT;
    by_Cur_Key :	BYTE;
    by_Attr :	BYTE;
    st_String :	STRING;
  END_VAR

  VAR
    us_TN_MENU_POPUP :	us_TN_MENU_POPUP;
    FB_TN_INPUT_MENU_POPUP :	TN_INPUT_MENU_POPUP;
    FB_TN_SC_WRITE :	TN_SC_WRITE;
    FB_FIX :	FIX;
    ELEMENT_COUNT :	ELEMENT_COUNT;
    ELEMENT_GET :	ELEMENT_GET;
  END_VAR

  VAR_IN_OUT
    Xus_TN_SCREEN :	us_TN_SCREEN;
    Xus_TN_INPUT_CONTROL_DATA :	us_TN_INPUT_CONTROL_DATA;
  END_VAR

  IF (Xus_TN_INPUT_CONTROL_DATA.bo_Focus = TRUE) THEN

    by_Cur_Key := Xus_TN_INPUT_CONTROL_DATA.by_Input_Exten_Code;

    IF (us_TN_MENU_POPUP.bo_Activ = FALSE) THEN
      us_TN_MENU_POPUP.by_Input_Exten_Code := BYTE#00;

      IF (by_Cur_Key = BYTE#13) THEN
        us_TN_MENU_POPUP.in_Y         := Xus_TN_INPUT_CONTROL_DATA.in_Y;
        us_TN_MENU_POPUP.in_X         := Xus_TN_INPUT_CONTROL_DATA.in_X;
        us_TN_MENU_POPUP.by_Attr_mF   := Xus_TN_INPUT_CONTROL_DATA.by_Attr_mF;
        us_TN_MENU_POPUP.by_Attr_oF   := Xus_TN_INPUT_CONTROL_DATA.by_Attr_oF;
        us_TN_MENU_POPUP.st_Menu_Text := Xus_TN_INPUT_CONTROL_DATA.st_Input_Data;
        us_TN_MENU_POPUP.bo_Create    := TRUE;
        us_TN_MENU_POPUP.in_Cur_Item  := INT#00;
      END_IF;

      IF (us_TN_MENU_POPUP.in_Cur_Item > INT#00) THEN
        Xus_TN_INPUT_CONTROL_DATA.in_selected      := us_TN_MENU_POPUP.in_Cur_Item;
        Xus_TN_INPUT_CONTROL_DATA.bo_Input_Entered := TRUE;
        Xus_TN_INPUT_CONTROL_DATA.bo_Update_Input  := TRUE;
        us_TN_MENU_POPUP.in_Cur_Item := INT#00;
      END_IF;

    ELSE
      us_TN_MENU_POPUP.by_Input_Exten_Code := by_Cur_Key;
    END_IF;

    FB_TN_INPUT_MENU_POPUP.Xus_TN_MENU_POPUP := us_TN_MENU_POPUP;
    FB_TN_INPUT_MENU_POPUP.Xus_TN_SCREEN     := Xus_TN_SCREEN;
    FB_TN_INPUT_MENU_POPUP();
    us_TN_MENU_POPUP := FB_TN_INPUT_MENU_POPUP.Xus_TN_MENU_POPUP;
    Xus_TN_SCREEN    := FB_TN_INPUT_MENU_POPUP.Xus_TN_SCREEN;

  END_IF;

  IF (Xus_TN_INPUT_CONTROL_DATA.bo_Update_Input = TRUE) OR (Xus_TN_INPUT_CONTROL_DATA.bo_Update_All = TRUE) THEN

    IF Xus_TN_INPUT_CONTROL_DATA.bo_Update_All = TRUE THEN

      IF (Xus_TN_INPUT_CONTROL_DATA.in_Title_X_Offset = INT#00) AND (Xus_TN_INPUT_CONTROL_DATA.in_Title_Y_Offset = INT#00) THEN
        FB_TN_SC_WRITE.Iin_Y := Xus_TN_INPUT_CONTROL_DATA.in_Y;
        FB_TN_SC_WRITE.Iin_X := Xus_TN_INPUT_CONTROL_DATA.in_X - LEN(Xus_TN_INPUT_CONTROL_DATA.st_Title_String);

      ELSE
        FB_TN_SC_WRITE.Iin_Y := Xus_TN_INPUT_CONTROL_DATA.in_Y + Xus_TN_INPUT_CONTROL_DATA.in_Title_Y_Offset;
        FB_TN_SC_WRITE.Iin_X := Xus_TN_INPUT_CONTROL_DATA.in_X + Xus_TN_INPUT_CONTROL_DATA.in_Title_X_Offset;

      END_IF;

      FB_TN_SC_WRITE.Iby_ATTR      := Xus_TN_INPUT_CONTROL_DATA.by_Title_Attr;
      FB_TN_SC_WRITE.Ist_STRING    := Xus_TN_INPUT_CONTROL_DATA.st_Title_String;
      FB_TN_SC_WRITE.Xus_TN_SCREEN := Xus_TN_SCREEN;
      FB_TN_SC_WRITE();
      Xus_TN_SCREEN := FB_TN_SC_WRITE.Xus_TN_SCREEN;

    END_IF;

    ELEMENT_COUNT(SEP:=BYTE#35,ELEMENT:=Xus_TN_INPUT_CONTROL_DATA.st_Input_Data);
    Xus_TN_INPUT_CONTROL_DATA.st_Input_Data:=ELEMENT_COUNT.ELEMENT;
    in_Element_Count:=ELEMENT_COUNT.ELEMENT_COUNT;

    IF in_Element_Count > INT#00 THEN

      Xus_TN_INPUT_CONTROL_DATA.in_selected:=LIMIT_INT(1,Xus_TN_INPUT_CONTROL_DATA.in_selected,in_Element_Count);

      in_index := Xus_TN_INPUT_CONTROL_DATA.in_selected;

      ELEMENT_GET(ELEMENT:=Xus_TN_INPUT_CONTROL_DATA.st_Input_Data,SEP:=BYTE#35,POS:=in_index-1);
      Xus_TN_INPUT_CONTROL_DATA.st_Input_Data:=ELEMENT_GET.ELEMENT;

      st_String:=ELEMENT_GET.ELEMENT_GET;

      FB_FIX.str:=st_String;
    FB_FIX.L:=LEN(Xus_TN_INPUT_CONTROL_DATA.st_Input_Mask);
    FB_FIX.C:=BYTE#32;
    FB_FIX.M:=Xus_TN_INPUT_CONTROL_DATA.in_Input_Option;
      FB_FIX();
      st_String:=FB_FIX.FIX;

      Xus_TN_INPUT_CONTROL_DATA.st_Input_String := st_String;

      IF Xus_TN_INPUT_CONTROL_DATA.bo_Focus = TRUE THEN
        by_Attr := Xus_TN_INPUT_CONTROL_DATA.by_Attr_mF;
      ELSE
        by_Attr := Xus_TN_INPUT_CONTROL_DATA.by_Attr_oF;
      END_IF;

      FB_TN_SC_WRITE.Iin_X         := Xus_TN_INPUT_CONTROL_DATA.in_X;
      FB_TN_SC_WRITE.Iin_Y         := Xus_TN_INPUT_CONTROL_DATA.in_Y;
      FB_TN_SC_WRITE.Iby_ATTR      := by_Attr;
      FB_TN_SC_WRITE.Ist_STRING    := st_String;
      FB_TN_SC_WRITE.Xus_TN_SCREEN := Xus_TN_SCREEN;
      FB_TN_SC_WRITE();
      Xus_TN_SCREEN := FB_TN_SC_WRITE.Xus_TN_SCREEN;

    END_IF;

    Xus_TN_INPUT_CONTROL_DATA.in_Cursor_X := Xus_TN_INPUT_CONTROL_DATA.in_X;
    Xus_TN_INPUT_CONTROL_DATA.in_Cursor_Y := Xus_TN_INPUT_CONTROL_DATA.in_Y;

    Xus_TN_INPUT_CONTROL_DATA.bo_Update_All   := FALSE;
    Xus_TN_INPUT_CONTROL_DATA.bo_Update_Input := FALSE;

  END_IF;

END_FUNCTION_BLOCK

(* ---- 676-RDM2.ST ---- *)
FUNCTION _REAL_TO_DWORD: DWORD
	VAR_INPUT
		X :	REAL;
	END_VAR

	IF REAL_TO_DWORD(0.5) = DWORD#1 THEN
		_REAL_TO_DWORD := REAL_TO_DWORD(x);
	ELSIF X > 0.0 THEN
		_REAL_TO_DWORD := REAL_TO_DWORD(x+0.5);
	ELSIF X < 0.0 THEN
		_REAL_TO_DWORD := REAL_TO_DWORD(x-0.5);
	ELSE
		_REAL_TO_DWORD := DWORD#0;
	END_IF;
END_FUNCTION

FUNCTION _DWORD_TO_REAL:REAL
	VAR_INPUT
		IN :	DWORD;
	END_VAR

	_DWORD_TO_REAL := UDINT_TO_REAL(DWORD_TO_UDINT(IN));

END_FUNCTION

FUNCTION _INT_TO_UDINT:UDINT
	VAR_INPUT
		IN :	INT;
	END_VAR

	_INT_TO_UDINT := DINT_TO_UDINT(INT_TO_DINT(IN));
END_FUNCTION

FUNCTION D_TRUNC : DINT
	VAR_INPUT
		x : REAL;
	END_VAR

	D_TRUNC := REAL_TO_DINT(X);
	IF X > 0.0 THEN
		IF DINT_TO_REAL(D_TRUNC) > X THEN D_TRUNC := D_TRUNC - DINT#1; END_IF;
	ELSE
		IF DINT_TO_REAL(D_TRUNC) < X THEN D_TRUNC := D_TRUNC + DINT#1; END_IF;
	END_IF;
END_FUNCTION

FUNCTION FRACT:REAL
	VAR_INPUT
		X :	REAL;
	END_VAR

	IF ABS(x) < 2.0E9 THEN
		FRACT := x - DINT_TO_REAL(D_TRUNC(x));
	ELSE
		FRACT := 0.0;
	END_IF;
END_FUNCTION

FUNCTION BIT_LOAD_DW:DWORD

	VAR_INPUT
		IN :	DWORD;
		VAL :	BOOL;
		POS :	INT;
	END_VAR

	IF val THEN
		BIT_LOAD_DW := in OR SHL(DWORD#1,pos);
	ELSE
		BIT_LOAD_DW := in AND (NOT SHL(DWORD#1,pos));
	END_IF;
END_FUNCTION

FUNCTION BIT_OF_DWORD : BOOL
	VAR_INPUT
		IN : DWORD;
		N : INT;
	END_VAR

	BIT_OF_DWORD := (SHR(in,N) AND 16#00000001) > 0;
END_FUNCTION

FUNCTION BIT_COUNT:INT
	VAR_INPUT
		IN :	DWORD;
	END_VAR

	VAR
		in_temp :	DWORD;
	END_VAR

	in_temp := IN;
	WHILE in_temp > DWORD#0 DO
		IF (in_temp AND DWORD#16#00000001) > DWORD#0 THEN Bit_Count := Bit_Count +1; END_IF;
		in_temp := SHR(in_temp,1);
	END_WHILE;
END_FUNCTION

FUNCTION_BLOCK T_PLC_MS_Block
	VAR_OUTPUT
		T_PLC_MS :	UDINT;
	END_VAR

	VAR_EXTERNAL
		PLC_TICKS_PER_SEC :	INT;
		PLC_SYS_TICK_CNT :	DINT;
	END_VAR

	VAR
		debug :	BOOL;(*Debug-Mode ON / OFF*)
		N :	INT;(*Debug-Faktor*)
		Offset :	UDINT;(*Debug-Offset*)
		temp :	DWORD := DWORD#1;(*Debug-Offset*)
		mode :	BOOL;(*modus*)
		faktor :	UDINT;(*Systemtakt-Faktor*)
		init :	BOOL;
		v_plc_ticks_per_sec :	UDINT;
		base :	UDINT := UDINT#1000;
	END_VAR

	IF init = FALSE THEN
		v_plc_ticks_per_sec := INT_TO_UDINT(PLC_TICKS_PER_SEC);
		IF v_plc_ticks_per_sec = UDINT#1024 THEN
			faktor := UDINT#1;
			mode := FALSE;
		ELSIF v_plc_ticks_per_sec > UDINT#0 THEN
			IF v_plc_ticks_per_sec <= base THEN
				faktor := base / v_plc_ticks_per_sec;
				mode := FALSE;
			ELSE
				faktor := v_plc_ticks_per_sec / base;
				mode := TRUE;
			END_IF;
		ELSE
			faktor := UDINT#1;
		END_IF;
		init := TRUE;
	END_IF;

	IF mode THEN
		T_PLC_MS := DINT_TO_UDINT(PLC_SYS_TICK_CNT) / faktor;
	ELSE
		T_PLC_MS := DINT_TO_UDINT(PLC_SYS_TICK_CNT) * faktor;
	END_IF;

	IF debug THEN
		T_PLC_MS := (DWORD_TO_UDINT(SHL(UDINT_TO_DWORD(T_PLC_MS),N) OR SHL(temp,N)) - UDINT#1) + Offset;
	END_IF;
END_FUNCTION_BLOCK

FUNCTION_BLOCK RDM_Block
	VAR_INPUT
		LAST :	REAL;
	END_VAR
	VAR_OUTPUT
		RDM :	REAL;
	END_VAR
	VAR
		T_PLC_MS :	T_PLC_MS_Block;
		tn :	DWORD;
		tc :	INT;
	END_VAR
	T_PLC_MS();
	tn := UDINT_TO_DWORD(T_PLC_MS.T_PLC_MS);
	tc := Bit_Count(tn);

	tn:=BIT_LOAD_DW(tn,BIT_OF_DWORD(tn,2),31); (* tn.31 := tn.2; *)
	tn:=BIT_LOAD_DW(tn,BIT_OF_DWORD(tn,5),30); (* tn.30 := tn.5; *)
	tn:=BIT_LOAD_DW(tn,BIT_OF_DWORD(tn,4),29); (* tn.29 := tn.4; *)
	tn:=BIT_LOAD_DW(tn,BIT_OF_DWORD(tn,1),28); (* tn.28 := tn.1; *)
	tn:=BIT_LOAD_DW(tn,BIT_OF_DWORD(tn,0),27); (* tn.27 := tn.0; *)
	tn:=BIT_LOAD_DW(tn,BIT_OF_DWORD(tn,7),26); (* tn.26 := tn.7; *)
	tn:=BIT_LOAD_DW(tn,BIT_OF_DWORD(tn,6),25); (* tn.25 := tn.6; *)
	tn:=BIT_LOAD_DW(tn,BIT_OF_DWORD(tn,3),24); (* tn.24 := tn.3; *)

	tn := ROL(tn,Bit_Count(tn)) OR DWORD#16#80000001;
	tn := UDINT_TO_DWORD(DWORD_TO_UDINT(tn) MOD UDINT#71474513 + _INT_TO_UDINT(tc) + UDINT#77);
	RDM := fract(_DWORD_TO_REAL(tn) / 10000000.0 * (2.71828182845904523536028747135266249 - LIMIT_REAL(0.0,last,1.0)));
END_FUNCTION_BLOCK

FUNCTION_BLOCK RDM2_Block
	VAR_INPUT
		LAST :	INT;
		LOW :	INT;
		HIGH :	INT;
	END_VAR

	VAR_OUTPUT
		RDM2 :	INT;
	END_VAR

	VAR
		rdm :	RDM_Block;
	END_VAR

	rdm(last:=fract(INT_TO_REAL(last) * 3.14159265358979323846264338327950288));
	RDM2 := TRUNC(rdm.RDM * INT_TO_REAL(high - low + 1)) + low;

END_FUNCTION_BLOCK

PROGRAM program0

	VAR
		LAST :	INT;
		LOW :	INT;
		HIGH :	INT;

        RDM2 :	INT;
		func_block : RDM2_Block;
	END_VAR
		func_block.LAST := LAST;
		func_block.LOW := LOW;
		func_block.HIGH := HIGH;
		func_block();
		RDM2 := func_block.RDM2;

END_PROGRAM

CONFIGURATION Config0

	VAR_GLOBAL
		PLC_TICKS_PER_SEC :	INT;
		PLC_SYS_TICK_CNT :	DINT;
	END_VAR

	RESOURCE Res0 ON PLC
		TASK task0(INTERVAL := T#20ms,PRIORITY := 0);
		PROGRAM instance0 WITH task0 : program0;
	END_RESOURCE

END_CONFIGURATION

(* ---- 677-GEN_RDM.ST ---- *)
FUNCTION D_TRUNC : DINT
  VAR_INPUT
    x : REAL;
  END_VAR

  D_TRUNC := REAL_TO_DINT(X);
  IF X > 0.0 THEN
  	IF DINT_TO_REAL(D_TRUNC) > X THEN D_TRUNC := D_TRUNC - DINT#1; END_IF;
  ELSE
  	IF DINT_TO_REAL(D_TRUNC) < X THEN D_TRUNC := D_TRUNC + DINT#1; END_IF;
  END_IF;
END_FUNCTION

FUNCTION BIT_COUNT:INT

	VAR_INPUT
		IN :	DWORD;
	END_VAR

	VAR
		in_temp :	DWORD;
	END_VAR

	in_temp := IN;
	WHILE in_temp > DWORD#0 DO
		IF (in_temp AND DWORD#16#00000001) > DWORD#0 THEN Bit_Count := Bit_Count +1; END_IF;
		in_temp := SHR(in_temp,1);
	END_WHILE;

END_FUNCTION

FUNCTION FRACT:REAL
	VAR_INPUT
		X :	REAL;
	END_VAR

	IF ABS(x) < 2.0E9 THEN
		FRACT := x - DINT_TO_REAL(D_TRUNC(x));
	ELSE
		FRACT := 0.0;
	END_IF;

END_FUNCTION

FUNCTION_BLOCK T_PLC_MS_block
	VAR_OUTPUT
		T_PLC_MS :	UDINT;
	END_VAR

	VAR_EXTERNAL
		PLC_TICKS_PER_SEC :	INT;
		PLC_SYS_TICK_CNT :	DINT;
	END_VAR

	VAR
		debug :	BOOL;(*Debug-Mode ON / OFF*)
		N :	INT;(*Debug-Faktor*)
		Offset :	UDINT;(*Debug-Offset*)
		temp :	DWORD := DWORD#1;(*Debug-Offset*)
		mode :	BOOL;(*modus*)
		faktor :	UDINT;(*Systemtakt-Faktor*)
		init :	BOOL;
		v_plc_ticks_per_sec :	UDINT;
		base :	UDINT := UDINT#1000;
	END_VAR

	IF init = FALSE THEN
		v_plc_ticks_per_sec := INT_TO_UDINT(PLC_TICKS_PER_SEC);
		IF v_plc_ticks_per_sec = UDINT#1024 THEN
			faktor := UDINT#1;
			mode := FALSE;
		ELSIF v_plc_ticks_per_sec > UDINT#0 THEN
			IF v_plc_ticks_per_sec <= base THEN
				faktor := base / v_plc_ticks_per_sec;
				mode := FALSE;
			ELSE
				faktor := v_plc_ticks_per_sec / base;
				mode := TRUE;
			END_IF;
		ELSE
			faktor := UDINT#1;
		END_IF;
		init := TRUE;
	END_IF;

	IF mode THEN
		T_PLC_MS := DINT_TO_UDINT(PLC_SYS_TICK_CNT) / faktor;
	ELSE
		T_PLC_MS := DINT_TO_UDINT(PLC_SYS_TICK_CNT) * faktor;
	END_IF;

	IF debug THEN
		T_PLC_MS := (DWORD_TO_UDINT(SHL(UDINT_TO_DWORD(T_PLC_MS),N) OR SHL(temp,N)) - UDINT#1) + Offset;
	END_IF;

END_FUNCTION_BLOCK

FUNCTION BIT_LOAD_DW:DWORD

	VAR_INPUT
		IN :	DWORD;
		VAL :	BOOL;
		POS :	INT;
	END_VAR

	IF val THEN
		BIT_LOAD_DW := in OR SHL(DWORD#1,pos);
	ELSE
		BIT_LOAD_DW := in AND (NOT SHL(DWORD#1,pos));
	END_IF;

END_FUNCTION

FUNCTION BIT_OF_DWORD : BOOL
  VAR_INPUT
    IN : DWORD;
    N : INT;
  END_VAR

  BIT_OF_DWORD := (SHR(in,N) AND 16#00000001) > 0;
  (* from OSCAT library; www.oscat.de  *)
END_FUNCTION

FUNCTION _INT_TO_UDINT:UDINT
	VAR_INPUT
		IN :	INT;
	END_VAR

	_INT_TO_UDINT := DINT_TO_UDINT(INT_TO_DINT(IN));
END_FUNCTION

FUNCTION _DWORD_TO_REAL:REAL
	VAR_INPUT
		IN :	DWORD;
	END_VAR

	_DWORD_TO_REAL := UDINT_TO_REAL(DWORD_TO_UDINT(IN));

END_FUNCTION

FUNCTION_BLOCK RDM_block
	VAR_INPUT
		LAST :	REAL;
	END_VAR
	VAR_OUTPUT
		RDM :	REAL;
	END_VAR
	VAR
		T_PLC_MS :	T_PLC_MS_block;
		tn :	DWORD;
		tc :	INT;
	END_VAR
	T_PLC_MS();
	tn := UDINT_TO_DWORD(T_PLC_MS.T_PLC_MS);
	tc := Bit_Count(tn);

	tn:=BIT_LOAD_DW(tn,BIT_OF_DWORD(tn,2),31); (* tn.31 := tn.2; *)
	tn:=BIT_LOAD_DW(tn,BIT_OF_DWORD(tn,5),30); (* tn.30 := tn.5; *)
	tn:=BIT_LOAD_DW(tn,BIT_OF_DWORD(tn,4),29); (* tn.29 := tn.4; *)
	tn:=BIT_LOAD_DW(tn,BIT_OF_DWORD(tn,1),28); (* tn.28 := tn.1; *)
	tn:=BIT_LOAD_DW(tn,BIT_OF_DWORD(tn,0),27); (* tn.27 := tn.0; *)
	tn:=BIT_LOAD_DW(tn,BIT_OF_DWORD(tn,7),26); (* tn.26 := tn.7; *)
	tn:=BIT_LOAD_DW(tn,BIT_OF_DWORD(tn,6),25); (* tn.25 := tn.6; *)
	tn:=BIT_LOAD_DW(tn,BIT_OF_DWORD(tn,3),24); (* tn.24 := tn.3; *)

	tn := ROL(tn,Bit_Count(tn)) OR DWORD#16#80000001;
	tn := UDINT_TO_DWORD(DWORD_TO_UDINT(tn) MOD UDINT#71474513 + _INT_TO_UDINT(tc) + UDINT#77);
	RDM := fract(_DWORD_TO_REAL(tn) / 10000000.0 * (2.71828182845904523536028747135266249 - LIMIT_REAL(0.0,last,1.0)));
END_FUNCTION_BLOCK

FUNCTION_BLOCK GEN_RDM_Block

	VAR_INPUT
		PT :	TIME;
		AM :	REAL := REAL#1.0;
		OS :	REAL;
	END_VAR

	VAR_OUTPUT
		Q :	BOOL;
		Out :	REAL;
	END_VAR

	VAR
		tx :	TIME;
		last :	TIME;
		init :	BOOL;
		T_PLC_MS :	T_PLC_MS_Block;
		FB_rdm :	RDM_block;
	END_VAR

	T_PLC_MS();
	tx:= UDINT_TO_TIME(T_PLC_MS.T_PLC_MS) - last;

	IF NOT init THEN
		init := TRUE;
		last := tx;
		tx := t#0s;
	END_IF;

	IF tx >= pt THEN
		last := last + pt;
		tx := tx - pt;

		FB_rdm(last:=0.0);
		out := am * (FB_rdm.RDM - 0.5) + os;
		q := TRUE;
	ELSE
		q := FALSE;
	END_IF;

END_FUNCTION_BLOCK

PROGRAM program0
  VAR
	PT :	TIME;
	AM :	REAL := REAL#1.0;
	OS :	REAL;
	Q :	BOOL;
	Out :	REAL;
	func_block : GEN_RDM_Block;
  END_VAR
	func_block.PT  :=PT;
	func_block.AM  :=AM;
	func_block.OS  :=OS;
	func_block();
	Q := func_block.Q;
	Out := func_block.Out;
END_PROGRAM

CONFIGURATION Config0
	VAR_GLOBAL
		PLC_TICKS_PER_SEC :	INT;
		PLC_SYS_TICK_CNT :	DINT;
	END_VAR
	RESOURCE Res0 ON PLC
		TASK task0(INTERVAL := T#20ms,PRIORITY := 0);
		PROGRAM instance0 WITH task0 : program0;
	END_RESOURCE
END_CONFIGURATION

(* ---- 678-RTC_2.ST ---- *)
FUNCTION _INT_TO_UDINT:UDINT
	VAR_INPUT
		IN :	INT;
	END_VAR

	_INT_TO_UDINT := DINT_TO_UDINT(INT_TO_DINT(IN));
END_FUNCTION

FUNCTION SET_DATE:UDINT

	VAR_INPUT
		YEAR :	INT;
		MONTH :	INT;
		DAY :	INT;
	END_VAR

	VAR
		count :	INT;
	END_VAR

	IF month > 2 THEN
		count := (month - 1) * 30;
		IF month > 7 THEN
			count := count + DWORD_TO_INT(SHR(DINT_TO_DWORD(INT_TO_DINT(month) - INT_TO_DINT(3)),1));
		ELSE
			count := count + DWORD_TO_INT(SHR(DINT_TO_DWORD(INT_TO_DINT(month) - INT_TO_DINT(4)),1));
		END_IF;
		IF SHL(INT_TO_WORD(year),14) = WORD#0 THEN
			count := count + 1;
		END_IF;
	ELSE
		count := (month - 1) * 31;
	END_IF;
	SET_DATE := (_INT_TO_UDINT(count + day - 1) + DWORD_TO_UDINT(SHR(UDINT_TO_DWORD(_INT_TO_UDINT(year) * UDINT#1461 - UDINT#2878169), 2))) * UDINT#86400;

END_FUNCTION

FUNCTION SET_DT:UDINT
	VAR_INPUT
		YEAR :	INT;
		MONTH :	INT;
		DAY :	INT;
		HOUR :	INT;
		MINUTE :	INT;
		SECOND :	INT;
	END_VAR

	SET_DT := SET_DATE(YEAR, MONTH, DAY) + _INT_TO_UDINT(SECOND) + _INT_TO_UDINT(MINUTE) * UDINT#60 + _INT_TO_UDINT(HOUR) * UDINT#3600;
END_FUNCTION

FUNCTION DT_TO_DATE2:UDINT

	VAR_INPUT
		IN :	UDINT;
	END_VAR

	DT_TO_DATE2 := (IN / UDINT#86400) * UDINT#86400;

END_FUNCTION

FUNCTION YEAR_OF_DATE:INT
	VAR_INPUT
		IDATE :	UDINT;
	END_VAR

	YEAR_OF_DATE := UDINT_TO_INT((idate+UDINT#43200) / UDINT#31557600 + UDINT#1970);
END_FUNCTION

FUNCTION DST:BOOL
	VAR_INPUT
		UTC :	UDINT;
	END_VAR

	VAR
		yr :	INT;
		yr4 :	UDINT;
		ltc :	UDINT;
		idate :	UDINT;
	END_VAR

	yr := YEAR_OF_DATE(DT_TO_DATE2(UTC));
	ltc := UTC;
	idate := SET_DT(yr, 3, 31, 1, 0, 0);
	yr4 := DWORD_TO_UDINT(SHR(INT_TO_DWORD(5 * yr), 2)) + UDINT#1;
	DST := (idate - ((yr4 + UDINT#3) MOD UDINT#7) * UDINT#86400 <= ltc) AND (idate + (UDINT#214 - (yr4) MOD UDINT#7) * UDINT#86400 > ltc);

END_FUNCTION

FUNCTION_BLOCK T_PLC_MS_Block
	VAR_OUTPUT
		T_PLC_MS :	UDINT;
	END_VAR

	VAR_EXTERNAL
		PLC_TICKS_PER_SEC :	INT;
		PLC_SYS_TICK_CNT :	DINT;
	END_VAR

	VAR
		debug :	BOOL;(*Debug-Mode ON / OFF*)
		N :	INT;(*Debug-Faktor*)
		Offset :	UDINT;(*Debug-Offset*)
		temp :	DWORD := DWORD#1;(*Debug-Offset*)
		mode :	BOOL;(*modus*)
		faktor :	UDINT;(*Systemtakt-Faktor*)
		init :	BOOL;
		v_plc_ticks_per_sec :	UDINT;
		base :	UDINT := UDINT#1000;
	END_VAR

	IF init = FALSE THEN
		v_plc_ticks_per_sec := INT_TO_UDINT(PLC_TICKS_PER_SEC);
		IF v_plc_ticks_per_sec = UDINT#1024 THEN
			faktor := UDINT#1;
			mode := FALSE;
		ELSIF v_plc_ticks_per_sec > UDINT#0 THEN
			IF v_plc_ticks_per_sec <= base THEN
				faktor := base / v_plc_ticks_per_sec;
				mode := FALSE;
			ELSE
				faktor := v_plc_ticks_per_sec / base;
				mode := TRUE;
			END_IF;
		ELSE
			faktor := UDINT#1;
		END_IF;
		init := TRUE;
	END_IF;

	IF mode THEN
		T_PLC_MS := DINT_TO_UDINT(PLC_SYS_TICK_CNT) / faktor;
	ELSE
		T_PLC_MS := DINT_TO_UDINT(PLC_SYS_TICK_CNT) * faktor;
	END_IF;

	IF debug THEN
		T_PLC_MS := (DWORD_TO_UDINT(SHL(UDINT_TO_DWORD(T_PLC_MS),N) OR SHL(temp,N)) - UDINT#1) + Offset;
	END_IF;
END_FUNCTION_BLOCK

FUNCTION_BLOCK RTC_MS_Block

	VAR_INPUT
		SET :	BOOL;
		SDT :	UDINT;
		SMS :	INT;
	END_VAR

	VAR_OUTPUT
		XDT :	UDINT;
		XMS :	INT;
	END_VAR

	VAR
		init :	BOOL;
		last :	UDINT;
		tx :	UDINT;
		T_PLC_MS :	T_PLC_MS_Block;
	END_VAR

	T_PLC_MS();
	tx:= T_PLC_MS.T_PLC_MS;

	IF set OR NOT init THEN
		(* clock needs to be set when set is true or after power up *)
		init := TRUE;
		xdt := SDT;
		XMS := SMS;
	ELSE
		XMS := XMS + UDINT_TO_INT(tx - last);
		(* check if one second has expired *)
		IF XMS > 999 THEN
			XDT := XDT + UDINT#1; (* add one second *)
			XMS := XMS - 1000;
		END_IF;
	END_IF;
	last := tx;

END_FUNCTION_BLOCK

FUNCTION_BLOCK RTC_2_Block

	VAR_INPUT
		SET :	BOOL;
		SDT :	UDINT;
		SMS :	INT;
		DEN :	BOOL;
		OFS :	INT;
	END_VAR

	VAR_OUTPUT
		UDT :	UDINT;
		LDT :	UDINT;
		DSO :	BOOL;
		XMS :	INT;
	END_VAR

	VAR
		RT :	RTC_MS_Block;
	END_VAR

	RT(SET := SET, SDT := SDT, SMS := SMS);
	UDT := rt.xdt;
	XMS := rt.XMS;

	dso := DST(udt) AND DEN;

	LDT := UDT + _INT_TO_UDINT(ofs + BOOL_TO_INT(DSO) * 60) * UDINT#60;

END_FUNCTION_BLOCK

PROGRAM program0

	VAR
		SET :	BOOL;
		SDT :	UDINT;
		SMS :	INT;
		DEN :	BOOL;
		OFS :	INT;
		UDT :	UDINT;
		LDT :	UDINT;
		DSO :	BOOL;
		XMS :	INT;
		func_block : RTC_2_Block;
  	END_VAR
	func_block.SET  :=	SET;
	func_block.SDT  :=	SDT;
	func_block.SMS  :=	SMS;
	func_block.DEN  :=	DEN;
	func_block.OFS  :=	OFS;
	func_block();
	UDT := func_block.UDT;
	LDT := func_block.LDT;
	DSO := func_block.DSO;
	XMS := func_block.XMS;

END_PROGRAM

CONFIGURATION Config0

	VAR_GLOBAL
		PLC_TICKS_PER_SEC :	INT;
		PLC_SYS_TICK_CNT :	DINT;
	END_VAR

	RESOURCE Res0 ON PLC
		TASK task0(INTERVAL := T#20ms,PRIORITY := 0);
		PROGRAM instance0 WITH task0 : program0;
	END_RESOURCE

END_CONFIGURATION

(* ---- 679-BLIND_ACTUATOR.ST ---- *)
FUNCTION_BLOCK INTERLOCK_Block

	VAR_INPUT
		I1 :	BOOL;
		I2 :	BOOL;
		TL :	TIME;
	END_VAR

	VAR_OUTPUT
		Q1 :	BOOL;
		Q2 :	BOOL;
	END_VAR

	VAR
		T1 :	TOF;
		T2 :	TOF;
	END_VAR

	T1(IN := I1, PT := TL);
	T2(IN := I2, PT := TL);

	Q1 := I1 AND NOT t2.Q;
	Q2 := I2 AND NOT t1.Q;

END_FUNCTION_BLOCK

FUNCTION TIME_TO_UDINT2:UDINT
	VAR_INPUT
		X :	TIME;
	END_VAR

	TIME_TO_UDINT2 := DINT_TO_UDINT(TIME_TO_DINT(X));
END_FUNCTION

FUNCTION_BLOCK T_PLC_MS_block
	VAR_OUTPUT
		T_PLC_MS :	UDINT;
	END_VAR

	VAR_EXTERNAL
		PLC_TICKS_PER_SEC :	INT;
		PLC_SYS_TICK_CNT :	DINT;
	END_VAR

	VAR
		debug :	BOOL;(*Debug-Mode ON / OFF*)
		N :	INT;(*Debug-Faktor*)
		Offset :	UDINT;(*Debug-Offset*)
		temp :	DWORD := DWORD#1;(*Debug-Offset*)
		mode :	BOOL;(*modus*)
		faktor :	UDINT;(*Systemtakt-Faktor*)
		init :	BOOL;
		v_plc_ticks_per_sec :	UDINT;
		base :	UDINT := UDINT#1000;
	END_VAR

	IF init = FALSE THEN
		v_plc_ticks_per_sec := INT_TO_UDINT(PLC_TICKS_PER_SEC);
		IF v_plc_ticks_per_sec = UDINT#1024 THEN
			faktor := UDINT#1;
			mode := FALSE;
		ELSIF v_plc_ticks_per_sec > UDINT#0 THEN
			IF v_plc_ticks_per_sec <= base THEN
				faktor := base / v_plc_ticks_per_sec;
				mode := FALSE;
			ELSE
				faktor := v_plc_ticks_per_sec / base;
				mode := TRUE;
			END_IF;
		ELSE
			faktor := UDINT#1;
		END_IF;
		init := TRUE;
	END_IF;

	IF mode THEN
		T_PLC_MS := DINT_TO_UDINT(PLC_SYS_TICK_CNT) / faktor;
	ELSE
		T_PLC_MS := DINT_TO_UDINT(PLC_SYS_TICK_CNT) * faktor;
	END_IF;

	IF debug THEN
		T_PLC_MS := (DWORD_TO_UDINT(SHL(UDINT_TO_DWORD(T_PLC_MS),N) OR SHL(temp,N)) - UDINT#1) + Offset;
	END_IF;
END_FUNCTION_BLOCK

FUNCTION FRMP_B:BYTE
	VAR_INPUT
		START :	BYTE;
		DIR :	BOOL;
		TD :	TIME;
		TR :	TIME;
	END_VAR

	IF TD < TR THEN
		FRMP_B := MIN(UDINT_TO_BYTE(DWORD_TO_UDINT(SHL(TIME_TO_DWORD(TD), 8)) / TIME_TO_UDINT2(TR)), SEL(DIR, START, USINT_TO_BYTE(USINT#255 - BYTE_TO_USINT(START))));
		IF DIR THEN
			FRMP_B := USINT_TO_BYTE(BYTE_TO_USINT(START) + BYTE_TO_USINT(FRMP_B));
		ELSE
			FRMP_B := USINT_TO_BYTE(BYTE_TO_USINT(START) - BYTE_TO_USINT(FRMP_B));
		END_IF;
	ELSE
		FRMP_B := SEL(DIR, BYTE#0, BYTE#255);
	END_IF;
END_FUNCTION

FUNCTION_BLOCK _RMP_B
	VAR_INPUT
		DIR :	BOOL;
		E :	BOOL := TRUE;
		TR :	TIME;
	END_VAR

	VAR_IN_OUT
		RMP :	BYTE;
	END_VAR

	VAR
		T_PLC_MS :	T_PLC_MS_block;
		tx :	TIME;
		tl :	TIME;
		tn :	TIME;
		init :	BOOL;
		last_dir :	BOOL;
		start :	BYTE;
	END_VAR

	T_PLC_MS();
	tx := UDINT_TO_TIME(T_PLC_MS.T_PLC_MS);

	IF E AND init AND (dir = last_dir) AND (RMP <> SEL(DIR, BYTE#0, BYTE#255)) AND TR = tn THEN
		RMP := FRMP_B(start, DIR, tx - tl, TR);
	ELSE
		init := TRUE;
		tl := tx;
		tn := tr;
		start := RMP;
	END_IF;
	last_dir := dir;
END_FUNCTION_BLOCK

FUNCTION_BLOCK RMP_B_Block

	VAR_INPUT
		SET :	BOOL;
		PT :	TIME;
		E :	BOOL := TRUE;
		UP :	BOOL := TRUE;
		RST :	BOOL;
	END_VAR

	VAR_OUTPUT
		OUT :	BYTE;
		BUSY :	BOOL;
		HIGH :	BOOL;
		LOW :	BOOL;
	END_VAR

	VAR
		rmp :	_RMP_B;
	END_VAR

	rmp(dir := UP, E := E, TR := PT, RMP := out);
	out := rmp.RMP;

	IF RST THEN
		out := BYTE#0;
	ELSIF SET THEN
		out := BYTE#255;
	END_IF;

low := out = BYTE#0;
high := out = BYTE#255;
busy := NOT (low OR high) AND E;

END_FUNCTION_BLOCK

FUNCTION_BLOCK BLIND_ACTUATOR_Block

	VAR_INPUT
		UP :	BOOL;
		DN :	BOOL;
		S_IN :	BYTE;
		T_UD :	TIME := T#10s;
		T_ANGLE :	TIME := T#3s;
		T_LOCKOUT :	TIME := t#100ms;
	END_VAR

	VAR_OUTPUT
		POS :	BYTE;
		ANG :	BYTE;
		QU :	BOOL;
		QD :	BOOL;
		STATUS :	BYTE;
	END_VAR

	VAR
		position :	RMP_B_Block;
		angle :	RMP_B_Block;
		lock :	INTERLOCK_Block;
	END_VAR

	lock(i1 := UP, I2 := DN, TL := T_lockout);

	angle(e := lock.Q1 OR lock.Q2, UP := lock.Q1, PT := T_Angle);
	position(e := lock.Q1 AND angle.high OR lock.Q2 AND angle.low, up := lock.Q1, PT := T_UD);

	pos := position.Out;
	ang := angle.Out;

	QU := lock.Q1;
	QD := lock.Q2;

	IF UP AND DN THEN
		status := BYTE#1;
	ELSIF UP THEN
		status := BYTE#121;
	ELSIF DN THEN
		status := BYTE#122;
	ELSE
		status := S_IN;
	END_IF;

END_FUNCTION_BLOCK

PROGRAM program0
	VAR
		UP :	BOOL;
		DN :	BOOL;
		S_IN :	BYTE;
		T_UD :	TIME := T#10s;
		T_ANGLE :	TIME := T#3s;
		T_LOCKOUT :	TIME := t#100ms;
		POS :	BYTE;
		ANG :	BYTE;
		QU :	BOOL;
		QD :	BOOL;
		func_block : BLIND_ACTUATOR_Block;
	END_VAR
	func_block.UP := UP;
	func_block.DN := DN;
	func_block.S_IN := S_IN ;
	func_block.T_UD := T_UD;
	func_block.T_ANGLE := T_ANGLE;
	func_block.T_LOCKOUT := T_LOCKOUT;
	func_block();
	POS  := func_block.POS;
	ANG  := func_block.ANG;
	QU  := func_block.QU;
	QD  := func_block.QD;
END_PROGRAM

CONFIGURATION Config0
	VAR_GLOBAL
		PLC_TICKS_PER_SEC :	INT;
		PLC_SYS_TICK_CNT :	DINT;
	END_VAR
  	RESOURCE Res0 ON PLC
    	TASK task0(INTERVAL := T#20ms,PRIORITY := 0);
    	PROGRAM instance0 WITH task0 : program0;
  	END_RESOURCE
END_CONFIGURATION

(* ---- 680-RDMDW.ST ---- *)
FUNCTION _REAL_TO_DWORD: DWORD
	VAR_INPUT
		X :	REAL;
	END_VAR

	IF REAL_TO_DWORD(0.5) = DWORD#1 THEN
		_REAL_TO_DWORD := REAL_TO_DWORD(x);
	ELSIF X > 0.0 THEN
		_REAL_TO_DWORD := REAL_TO_DWORD(x+0.5);
	ELSIF X < 0.0 THEN
		_REAL_TO_DWORD := REAL_TO_DWORD(x-0.5);
	ELSE
		_REAL_TO_DWORD := DWORD#0;
	END_IF;
END_FUNCTION

FUNCTION _DWORD_TO_REAL:REAL
	VAR_INPUT
		IN :	DWORD;
	END_VAR

	_DWORD_TO_REAL := UDINT_TO_REAL(DWORD_TO_UDINT(IN));

END_FUNCTION

FUNCTION _INT_TO_UDINT:UDINT
	VAR_INPUT
		IN :	INT;
	END_VAR

	_INT_TO_UDINT := DINT_TO_UDINT(INT_TO_DINT(IN));
END_FUNCTION

FUNCTION D_TRUNC : DINT
	VAR_INPUT
		x : REAL;
	END_VAR

	D_TRUNC := REAL_TO_DINT(X);
	IF X > 0.0 THEN
		IF DINT_TO_REAL(D_TRUNC) > X THEN D_TRUNC := D_TRUNC - DINT#1; END_IF;
	ELSE
		IF DINT_TO_REAL(D_TRUNC) < X THEN D_TRUNC := D_TRUNC + DINT#1; END_IF;
	END_IF;
END_FUNCTION

FUNCTION FRACT:REAL
	VAR_INPUT
		X :	REAL;
	END_VAR

	IF ABS(x) < 2.0E9 THEN
		FRACT := x - DINT_TO_REAL(D_TRUNC(x));
	ELSE
		FRACT := 0.0;
	END_IF;
END_FUNCTION

FUNCTION BIT_LOAD_DW:DWORD

	VAR_INPUT
		IN :	DWORD;
		VAL :	BOOL;
		POS :	INT;
	END_VAR

	IF val THEN
		BIT_LOAD_DW := in OR SHL(DWORD#1,pos);
	ELSE
		BIT_LOAD_DW := in AND (NOT SHL(DWORD#1,pos));
	END_IF;
END_FUNCTION

FUNCTION BIT_OF_DWORD : BOOL
	VAR_INPUT
		IN : DWORD;
		N : INT;
	END_VAR

	BIT_OF_DWORD := (SHR(in,N) AND 16#00000001) > 0;
END_FUNCTION

FUNCTION BIT_COUNT:INT
	VAR_INPUT
		IN :	DWORD;
	END_VAR

	VAR
		in_temp :	DWORD;
	END_VAR

	in_temp := IN;
	WHILE in_temp > DWORD#0 DO
		IF (in_temp AND DWORD#16#00000001) > DWORD#0 THEN Bit_Count := Bit_Count +1; END_IF;
		in_temp := SHR(in_temp,1);
	END_WHILE;
END_FUNCTION

FUNCTION_BLOCK T_PLC_MS_Block
	VAR_OUTPUT
		T_PLC_MS :	UDINT;
	END_VAR

	VAR_EXTERNAL
		PLC_TICKS_PER_SEC :	INT;
		PLC_SYS_TICK_CNT :	DINT;
	END_VAR

	VAR
		debug :	BOOL;(*Debug-Mode ON / OFF*)
		N :	INT;(*Debug-Faktor*)
		Offset :	UDINT;(*Debug-Offset*)
		temp :	DWORD := DWORD#1;(*Debug-Offset*)
		mode :	BOOL;(*modus*)
		faktor :	UDINT;(*Systemtakt-Faktor*)
		init :	BOOL;
		v_plc_ticks_per_sec :	UDINT;
		base :	UDINT := UDINT#1000;
	END_VAR

	IF init = FALSE THEN
		v_plc_ticks_per_sec := INT_TO_UDINT(PLC_TICKS_PER_SEC);
		IF v_plc_ticks_per_sec = UDINT#1024 THEN
			faktor := UDINT#1;
			mode := FALSE;
		ELSIF v_plc_ticks_per_sec > UDINT#0 THEN
			IF v_plc_ticks_per_sec <= base THEN
				faktor := base / v_plc_ticks_per_sec;
				mode := FALSE;
			ELSE
				faktor := v_plc_ticks_per_sec / base;
				mode := TRUE;
			END_IF;
		ELSE
			faktor := UDINT#1;
		END_IF;
		init := TRUE;
	END_IF;

	IF mode THEN
		T_PLC_MS := DINT_TO_UDINT(PLC_SYS_TICK_CNT) / faktor;
	ELSE
		T_PLC_MS := DINT_TO_UDINT(PLC_SYS_TICK_CNT) * faktor;
	END_IF;

	IF debug THEN
		T_PLC_MS := (DWORD_TO_UDINT(SHL(UDINT_TO_DWORD(T_PLC_MS),N) OR SHL(temp,N)) - UDINT#1) + Offset;
	END_IF;
END_FUNCTION_BLOCK

FUNCTION_BLOCK RDM_Block
	VAR_INPUT
		LAST :	REAL;
	END_VAR
	VAR_OUTPUT
		RDM :	REAL;
	END_VAR
	VAR
		T_PLC_MS :	T_PLC_MS_Block;
		tn :	DWORD;
		tc :	INT;
	END_VAR
	T_PLC_MS();
	tn := UDINT_TO_DWORD(T_PLC_MS.T_PLC_MS);
	tc := Bit_Count(tn);

	tn:=BIT_LOAD_DW(tn,BIT_OF_DWORD(tn,2),31); (* tn.31 := tn.2; *)
	tn:=BIT_LOAD_DW(tn,BIT_OF_DWORD(tn,5),30); (* tn.30 := tn.5; *)
	tn:=BIT_LOAD_DW(tn,BIT_OF_DWORD(tn,4),29); (* tn.29 := tn.4; *)
	tn:=BIT_LOAD_DW(tn,BIT_OF_DWORD(tn,1),28); (* tn.28 := tn.1; *)
	tn:=BIT_LOAD_DW(tn,BIT_OF_DWORD(tn,0),27); (* tn.27 := tn.0; *)
	tn:=BIT_LOAD_DW(tn,BIT_OF_DWORD(tn,7),26); (* tn.26 := tn.7; *)
	tn:=BIT_LOAD_DW(tn,BIT_OF_DWORD(tn,6),25); (* tn.25 := tn.6; *)
	tn:=BIT_LOAD_DW(tn,BIT_OF_DWORD(tn,3),24); (* tn.24 := tn.3; *)

	tn := ROL(tn,Bit_Count(tn)) OR DWORD#16#80000001;
	tn := UDINT_TO_DWORD(DWORD_TO_UDINT(tn) MOD UDINT#71474513 + _INT_TO_UDINT(tc) + UDINT#77);
	RDM := fract(_DWORD_TO_REAL(tn) / 10000000.0 * (2.71828182845904523536028747135266249 - LIMIT_REAL(0.0,last,1.0)));
END_FUNCTION_BLOCK

FUNCTION_BLOCK RDMDW_Block

	VAR_INPUT
		LAST :	DWORD;
	END_VAR

	VAR_OUTPUT
		RDMDW :	DWORD;
	END_VAR

	VAR
		RX :	REAL;
		M :	REAL;
		rdm :	RDM_Block;
	END_VAR

	M := INT_TO_REAL(BIT_COUNT(last));
	rdm(last:=FRACT(M*3.14159265358979323846264338327950288));
	RX:=rdm.RDM;
	RDMDW := SHL(_REAL_TO_DWORD(rx*65535.0),16);

	rdm(last:=FRACT(M*2.71828182845904523536028747135266249));
	RX:=rdm.RDM;
	RDMDW := RDMDW OR (_REAL_TO_DWORD(rx*65535.0) AND DWORD#16#0000FFFF);

END_FUNCTION_BLOCK

PROGRAM program0

	VAR
		LAST :	DWORD;

        RDMDW :	DWORD;
		func_block : RDMDW_Block;
	END_VAR
		func_block.LAST := LAST;
		func_block();
		RDMDW := func_block.RDMDW;

END_PROGRAM

CONFIGURATION Config0

	VAR_GLOBAL
		PLC_TICKS_PER_SEC :	INT;
		PLC_SYS_TICK_CNT :	DINT;
	END_VAR

	RESOURCE Res0 ON PLC
		TASK task0(INTERVAL := T#20ms,PRIORITY := 0);
		PROGRAM instance0 WITH task0 : program0;
	END_RESOURCE

END_CONFIGURATION

(* ---- 681-SHA1_STR.ST ---- *)
TYPE
  oscat_aB0_19	: ARRAY [0..19]	OF BYTE;
  oscat_aB0_63	: ARRAY [0..63]	OF BYTE;
  oscat_aDW0_4	: ARRAY [0..4] 	OF DWORD;
  oscat_sDW0_79	: ARRAY [0..79] OF DWORD;
oscat_STRING250             : STRING;
END_TYPE

FUNCTION DWORD_OF_BYTE:DWORD
	VAR_INPUT
		B3 :	BYTE;
		B2 :	BYTE;
		B1 :	BYTE;
		B0 :	BYTE;
	END_VAR

	DWORD_OF_BYTE := SHL(SHL(SHL(BYTE_TO_DWORD(B3),8) OR BYTE_TO_DWORD(B2),8) OR BYTE_TO_DWORD(B1),8) OR BYTE_TO_DWORD(B0);

END_FUNCTION

FUNCTION_BLOCK SHA1_STREAM_Block

	VAR_IN_OUT
		MODE :	INT;
		BUF :	oscat_aB0_63;
		SHA1 :	oscat_aB0_19;
		SIZE :	UDINT;
	END_VAR

	VAR_OUTPUT
		POS :	UDINT;
	END_VAR

	VAR
		hash :	oscat_aDW0_4;
		end :	UDINT;
		block :	UDINT;
		pad_1 :	BOOL;
		w :	oscat_sDW0_79;
		n :	INT;
		n1 :	INT;
		n2 :	INT;
		n3 :	INT;
		n4 :	INT;
		a :	DWORD;
		b :	DWORD;
		c :	DWORD;
		d :	DWORD;
		e :	DWORD;
		f :	DWORD;
		k :	DWORD;
		x :	DWORD;
	END_VAR

	CASE MODE OF

	1:
		hash[0] := DWORD#16#67452301;
		hash[1] := DWORD#16#EFCDAB89;
		hash[2] := DWORD#16#98BADCFE;
		hash[3] := DWORD#16#10325476;
		hash[4] := DWORD#16#C3D2E1F0;

		FOR n := 16 TO 79 DO
			w[n] := DWORD#0;
		END_FOR;

		block := DWORD_TO_UDINT(SHR(UDINT_TO_DWORD(SIZE),6)) + BOOL_TO_UDINT((UDINT_TO_BYTE(SIZE) AND BYTE#16#3F) > BYTE#55);

		pad_1 := FALSE;
		POS := UDINT#0;
		End := SIZE;
		SIZE := MIN(UDINT#64,End);
		MODE := 2;

	2:	FOR n := UDINT_TO_INT(SIZE) TO 63 DO
			BUF[n] := BYTE#0;
		END_FOR;

		IF SIZE < UDINT#64 AND NOT pad_1 THEN
			BUF[SIZE] := BYTE#2#1000_0000;
			pad_1 := TRUE;
		END_IF;

		POS := POS + SIZE;
		SIZE := MIN(UDINT#64,End - POS);

		n := 0;
		FOR n4 := 0 TO 15 DO
			n1 := n + 1;
			n2 := n + 2;
			n3 := n + 3;
			w[n4] := DWORD_OF_BYTE(BUF[n],BUF[n1],BUF[n2],BUF[n3]);
			n := n + 4;
		END_FOR;

		IF block = UDINT#0 THEN
			w[15] := SHL(UDINT_TO_DWORD(End),3);
			MODE := 3;
		ELSE
			block := block - UDINT#1;
		END_IF;

		FOR n := 16 TO 79 DO
			n1 := n - 3;
			n2 := n - 8;
			n3 := n - 14;
			n4 := n - 16;
			w[n] := ROL(w[n1] XOR w[n2] XOR w[n3] XOR w[n4],1);
		END_FOR;

		a := hash[0];
		b := hash[1];
		c := hash[2];
		d := hash[3];
		e := hash[4];

		FOR n := 0 TO 79 DO
			IF n <= 19 THEN
				f := (b AND c) OR (NOT(b) AND d);
				k := DWORD#16#5A827999;
			ELSIF n <= 39 THEN
				f := b XOR c XOR d;
				k := DWORD#16#6ED9EBA1;
			ELSIF n <= 59 THEN
				f := (b AND c) OR (b AND d) OR (c AND d);
				k := DWORD#16#8F1BBCDC;
			ELSE
				f := b XOR c XOR d;
				k := DWORD#16#CA62C1D6;
			END_IF;

			x := UDINT_TO_DWORD(DWORD_TO_UDINT(ROL(a,5)) + DWORD_TO_UDINT(f) + DWORD_TO_UDINT(e) + DWORD_TO_UDINT(k) + DWORD_TO_UDINT(w[n]));
			e := d;
			d := c;
			c := ROL(b,30);
			b := a;
			a := x;
		END_FOR;

		hash[0] := UDINT_TO_DWORD(DWORD_TO_UDINT(hash[0]) + DWORD_TO_UDINT(a));
		hash[1] := UDINT_TO_DWORD(DWORD_TO_UDINT(hash[1]) + DWORD_TO_UDINT(b));
		hash[2] := UDINT_TO_DWORD(DWORD_TO_UDINT(hash[2]) + DWORD_TO_UDINT(c));
		hash[3] := UDINT_TO_DWORD(DWORD_TO_UDINT(hash[3]) + DWORD_TO_UDINT(d));
		hash[4] := UDINT_TO_DWORD(DWORD_TO_UDINT(hash[4]) + DWORD_TO_UDINT(e));

	END_CASE;

	IF MODE = 3 THEN
		n2 := 0;
		FOR n := 0 TO 4 DO
			FOR n1 := 0 TO 3 DO
				hash[n] := ROL(hash[n],8);
				SHA1[n2] := DWORD_TO_BYTE(hash[n]);
				n2 := n2 + 1;
			END_FOR;
		END_FOR;
	END_IF;

END_FUNCTION_BLOCK

FUNCTION_BLOCK SHA1_STR_Block

	VAR_INPUT
		RUN :	BOOL;
	END_VAR

	VAR_OUTPUT
		DONE :	BOOL;
	END_VAR

	VAR_IN_OUT
		STR :	oscat_STRING250;
		SHA1 :	oscat_aB0_19;
	END_VAR

	VAR
		run_last :	BOOL;
		SHA1_STREAM :	SHA1_STREAM_Block;
		buf :	oscat_aB0_63;
		mode :	INT;
		size :	UDINT;
		pos :	UDINT;
		i :	INT;
		i2 :	INT;
		CODE :	CODE;
	END_VAR

	CASE mode OF
	0:
		IF RUN AND NOT run_last THEN
			DONE := FALSE;
			mode := 1;
			size := INT_TO_UDINT(LEN(STR));
		END_IF;

	2:
		IF size > UDINT#0 THEN
			i2 := 0;
			FOR i := 1 TO UDINT_TO_INT(SIZE) DO
				CODE(STR:=MID(STR,1,UDINT_TO_INT(POS) + i),POS:=1);
				buf[i2] := CODE.CODE;
				i2 := i2 + 1;
			END_FOR;
		END_IF;

	3:	DONE := TRUE;
		mode := 0;

	END_CASE;

	IF mode > 0 THEN
		SHA1_STREAM(MODE:=mode, BUF:=buf, SHA1:=SHA1, SIZE:=size);
		mode := SHA1_STREAM.MODE;
		buf := SHA1_STREAM.BUF;
		SHA1 := SHA1_STREAM.SHA1;
		size := SHA1_STREAM.SIZE;
		pos := SHA1_STREAM.POS;
	END_IF;

	run_last := RUN;

END_FUNCTION_BLOCK

PROGRAM program0
	VAR
		MODE :	INT;
		BUF :	oscat_aB0_63;
		SHA1 :	oscat_aB0_19;
		SIZE :	UDINT;
		POS :	UDINT;

		func_block : SHA1_STREAM_Block;
	END_VAR
	func_block.MODE := MODE;
	func_block.BUF := BUF;
	func_block.SHA1 := SHA1;
	func_block.SIZE := SIZE;

	func_block();
  	MODE  := func_block.MODE;
	BUF  := func_block.BUF;
	SHA1  := func_block.SHA1;
	SIZE  := func_block.SIZE;
	POS  := func_block.POS;
END_PROGRAM

CONFIGURATION Config0
	RESOURCE Res0 ON PLC
		TASK task0(INTERVAL := T#20ms,PRIORITY := 0);
		PROGRAM instance0 WITH task0 : program0;
	END_RESOURCE
END_CONFIGURATION

(* ---- 682-_RMP_NEXT.ST ---- *)
FUNCTION UDINT_TO_TIME2:TIME

	VAR_INPUT
		IN :	UDINT;
	END_VAR

	UDINT_TO_TIME2 := DINT_TO_TIME(UDINT_TO_DINT(IN));

END_FUNCTION

FUNCTION_BLOCK T_PLC_MS_block
	VAR_OUTPUT
		T_PLC_MS :	UDINT;
	END_VAR

	VAR_EXTERNAL
		PLC_TICKS_PER_SEC :	INT;
		PLC_SYS_TICK_CNT :	DINT;
	END_VAR

	VAR
		debug :	BOOL;(*Debug-Mode ON / OFF*)
		N :	INT;(*Debug-Faktor*)
		Offset :	UDINT;(*Debug-Offset*)
		temp :	DWORD := DWORD#1;(*Debug-Offset*)
		mode :	BOOL;(*modus*)
		faktor :	UDINT;(*Systemtakt-Faktor*)
		init :	BOOL;
		v_plc_ticks_per_sec :	UDINT;
		base :	UDINT := UDINT#1000;
	END_VAR

	IF init = FALSE THEN
		v_plc_ticks_per_sec := INT_TO_UDINT(PLC_TICKS_PER_SEC);
		IF v_plc_ticks_per_sec = UDINT#1024 THEN
			faktor := UDINT#1;
			mode := FALSE;
		ELSIF v_plc_ticks_per_sec > UDINT#0 THEN
			IF v_plc_ticks_per_sec <= base THEN
				faktor := base / v_plc_ticks_per_sec;
				mode := FALSE;
			ELSE
				faktor := v_plc_ticks_per_sec / base;
				mode := TRUE;
			END_IF;
		ELSE
			faktor := UDINT#1;
		END_IF;
		init := TRUE;
	END_IF;

	IF mode THEN
		T_PLC_MS := DINT_TO_UDINT(PLC_SYS_TICK_CNT) / faktor;
	ELSE
		T_PLC_MS := DINT_TO_UDINT(PLC_SYS_TICK_CNT) * faktor;
	END_IF;

	IF debug THEN
		T_PLC_MS := (DWORD_TO_UDINT(SHL(UDINT_TO_DWORD(T_PLC_MS),N) OR SHL(temp,N)) - UDINT#1) + Offset;
	END_IF;
END_FUNCTION_BLOCK

FUNCTION TIME_TO_UDINT2:UDINT
	VAR_INPUT
		X :	TIME;
	END_VAR

	TIME_TO_UDINT2 := DINT_TO_UDINT(TIME_TO_DINT(X));
END_FUNCTION

FUNCTION FRMP_B:BYTE
	VAR_INPUT
		START :	BYTE;
		DIR :	BOOL;
		TD :	TIME;
		TR :	TIME;
	END_VAR

	IF TD < TR THEN
		FRMP_B := MIN(UDINT_TO_BYTE(DWORD_TO_UDINT(SHL(TIME_TO_DWORD(TD), 8)) / TIME_TO_UDINT2(TR)), SEL(DIR, START, USINT_TO_BYTE(USINT#255 - BYTE_TO_USINT(START))));
		IF DIR THEN
			FRMP_B := USINT_TO_BYTE(BYTE_TO_USINT(START) + BYTE_TO_USINT(FRMP_B));
		ELSE
			FRMP_B := USINT_TO_BYTE(BYTE_TO_USINT(START) - BYTE_TO_USINT(FRMP_B));
		END_IF;
	ELSE
		FRMP_B := SEL(DIR, BYTE#0, BYTE#255);
	END_IF;
END_FUNCTION

FUNCTION_BLOCK _RMP_B
	VAR_INPUT
		DIR :	BOOL;
		E :	BOOL := TRUE;
		TR :	TIME;
	END_VAR

	VAR_IN_OUT
		RMP :	BYTE;
	END_VAR

	VAR
		T_PLC_MS :	T_PLC_MS_block;
		tx :	TIME;
		tl :	TIME;
		tn :	TIME;
		init :	BOOL;
		last_dir :	BOOL;
		start :	BYTE;
	END_VAR

	T_PLC_MS();
	tx := UDINT_TO_TIME(T_PLC_MS.T_PLC_MS);

	IF E AND init AND (dir = last_dir) AND (RMP <> SEL(DIR, BYTE#0, BYTE#255)) AND TR = tn THEN
		RMP := FRMP_B(start, DIR, tx - tl, TR);
	ELSE
		init := TRUE;
		tl := tx;
		tn := tr;
		start := RMP;
	END_IF;
	last_dir := dir;
END_FUNCTION_BLOCK

FUNCTION_BLOCK TREND_DW
	VAR_INPUT
		X :	DWORD;
	END_VAR
	VAR_OUTPUT
		Q :	BOOL;
		TU :	BOOL;
		TD :	BOOL;
		D :	DWORD;
	END_VAR

	VAR
		LAST_X :	DWORD;
	END_VAR

	IF X > last_X THEN
		TU := TRUE;
		TD := FALSE;
		D := UDINT_TO_DWORD(DWORD_TO_UDINT(X) - DWORD_TO_UDINT(last_X));
		Q := TRUE;
	ELSIF X < last_X THEN
		TD := TRUE;
		TU := FALSE;
		D := UDINT_TO_DWORD(DWORD_TO_UDINT(last_X) - DWORD_TO_UDINT(X));
		Q := FALSE;
	ELSE
		TU := FALSE;
		TD := FALSE;
		D := DWORD#0;
	END_IF;
	last_X := X;
END_FUNCTION_BLOCK

FUNCTION_BLOCK _RMP_NEXT
	VAR_INPUT
		E :	BOOL := TRUE;
		IN :	BYTE;
		TR :	TIME;
		TF :	TIME;
		TL :	TIME;
	END_VAR

	VAR_OUTPUT
		DIR :	BOOL;
		UP :	BOOL;
		DN :	BOOL;
	END_VAR

	VAR_IN_OUT
		OUT :	BYTE;
	END_VAR
	VAR
		rmx :	_RMP_B;
		dirx :	TREND_DW;
		t_lock :	TP;
		xen :	BOOL;
		xdir :	BOOL;
	END_VAR

	dirx(X := BYTE_TO_DWORD(in));

	t_lock(in := FALSE, pt := TL);

	IF dirx.TU AND (OUT < IN) THEN
		IF NOT xdir AND xen THEN t_lock(in := TRUE); END_IF;
		xen := TRUE;
		xdir := TRUE;
	ELSIF dirx.TD AND (OUT > IN) THEN
		IF xdir AND xen THEN t_lock(in := TRUE); END_IF;
		xen := TRUE;
		xdir := FALSE;
	ELSIF xen THEN
		IF (xdir AND (out >= in)) OR (NOT xdir AND (out <= in)) THEN
			xen := FALSE;
			IF tl > t#0s THEN t_lock(IN := TRUE); END_IF;
		END_IF;
	END_IF;

	IF NOT t_lock.Q AND xen THEN
		UP := XDIR;
		DIR := XDIR;
		DN := NOT XDIR;
	ELSE
		UP := FALSE;
		DN := FALSE;
	END_IF;

	rmx(rmp := OUT, E := E AND (UP OR DN) , dir := DIR, tr := SEL(dir, TF, TR));
	OUT := rmx.RMP;
END_FUNCTION_BLOCK

PROGRAM program0
	VAR
	    LocalVar1 : BOOL;
		LocalVar2 : BYTE;
		LocalVar3 : TIME;
		LocalVar4 : TIME;
		LocalVar5 : TIME;
		LocalVar6 : BOOL;
		LocalVar7 : BOOL;
		LocalVar8 : BOOL;
		LocalInOut : BYTE;
		func_block : _RMP_NEXT;
  	END_VAR
	func_block.E  := LocalVar1;
	func_block.IN := LocalVar2;
	func_block.TR := LocalVar3;
	func_block.TF := LocalVar4;
	func_block.TL := LocalVar5;
	func_block.OUT := LocalInOut;
	func_block();
	LocalInOut := func_block.OUT;
	LocalVar6 := func_block.DIR;
	LocalVar7 := func_block.UP;
	LocalVar8 := func_block.DN;
END_PROGRAM

CONFIGURATION Config0
	VAR_GLOBAL
		PLC_TICKS_PER_SEC :	INT;
		PLC_SYS_TICK_CNT :	DINT;
	END_VAR
  	RESOURCE Res0 ON PLC
    	TASK task0(INTERVAL := T#20ms,PRIORITY := 0);
    	PROGRAM instance0 WITH task0 : program0;
  	END_RESOURCE
END_CONFIGURATION
